  rq_init_comm_if_connected(9, "1")
  rq_init_comm_if_connected(2, "2")
  rq_init_comm_if_connected(3, "3")
  rq_init_comm_if_connected(4, "4")
  rq_print_connected_grippers()
  rq_gripper_communication_thread = run rq_gripper_communication()
  set_closed_norm(97.6470588235294, 1)
  set_open_norm(1.1764705882352942, 1)
  set_closed_mm(0.0, 1)
  set_open_mm(53.0, 1)
  set_closed_norm(100.0, 2)
  set_open_norm(0.0, 2)
  set_closed_mm(0.0, 2)
  set_open_mm(50.0, 2)
  set_closed_norm(100.0, 3)
  set_open_norm(0.0, 3)
  set_closed_mm(0.0, 3)
  set_open_mm(50.0, 3)
  set_closed_norm(100.0, 4)
  set_open_norm(0.0, 4)
  set_closed_mm(0.0, 4)
  set_open_mm(50.0, 4)
  rq_current_limit_enabled = False
  while(not rq_gripper_communication_thread_started):
      sync()
  end
  # end: URCap Installation Node
  # begin: URCap Installation Node
  #   Source: OPC UA, 2.0.2, Rocketfarm AS
  #   Type: OPC UA
  global opcua_daemon = rpc_factory("xmlrpc", "http://127.0.0.1:40409/RPC2")
  def opcua_client_connect(address):
  return opcua_daemon.client_connect(address)
  end
  def opcua_client_get_id(client_name):
  return opcua_daemon.client_get_id(client_name)
  end
  def opcua_client_try_connect(client_id):
  opcua_result = False
  if (opcua_daemon.client_connect(client_id)):
  sleep(0.01)
  opcua_result = opcua_daemon.client_is_connected(client_id)
  opcua_retry = 10
  while ( (not opcua_result) and (opcua_retry > 0) ):
  sleep(0.1)
  opcua_result = opcua_daemon.client_is_connected(client_id)
  opcua_retry = opcua_retry - 1
  end
  end
  return opcua_result
  end
  def opcua_client_disconnect(client_id):
  return opcua_daemon.client_disconnect(client_id)
  end
  def opcua_client_is_connected(client_id):
  return opcua_daemon.client_is_connected(client_id)
  end
  def opcua_client_read_byid(client_id, namespace_id, variable_id):
  return opcua_daemon.client_read_variable_by_id(client_id, namespace_id, variable_id)
  end
  def opcua_client_read_byname(client_id, namespace_id, variable_name):
  return opcua_daemon.client_read_variable_by_name(client_id, namespace_id, variable_name)
  end
  def opcua_client_write_byid(client_id, namespace_id, variable_id, variable_value):
  return opcua_daemon.client_write_variable_by_id(client_id, namespace_id, variable_id, variable_value)
  end
  def opcua_client_write_byname(client_id, namespace_id, variable_name, variable_value):
  return opcua_daemon.client_write_variable_by_name(client_id, namespace_id, variable_name, variable_value)
  end
  def opcua_client_last_error(client_id):
  return opcua_daemon.client_get_last_error(client_id)
  end
  def opcua_server_read_byname(variable_name):
  return opcua_daemon.server_read_variable_by_name(variable_name)
  end
  def opcua_server_write_byname(variable_name, variable_value):
  return opcua_daemon.server_write_variable_by_name(variable_name, variable_value)
  end
  def opcua_server_last_error():
  return opcua_daemon.server_get_last_error()
  end
  def opcua_error_to_string(errorCode):
  return opcua_daemon.error_code_to_string(errorCode)
  end
  # end: URCap Installation Node
  step_count_7f95097d_1581_4d0e_9124_3b7fc3d01574 = 0.0
  thread Step_Counter_Thread_7db62caa_18b4_480e_a8f7_ee898fbd2f33():
    while (True):
      step_count_7f95097d_1581_4d0e_9124_3b7fc3d01574 = step_count_7f95097d_1581_4d0e_9124_3b7fc3d01574 + 1.0
      sync()
    end
  end
  run Step_Counter_Thread_7db62caa_18b4_480e_a8f7_ee898fbd2f33()
  global AMR_Position=struct(position_identifier=0, x1=0, x2=0, y1=0, y2=0, theta1=0, theta2=0)
  global CAM_Pose=p[0,0,0,0,0,0]
  global CAM_Relation=""
  global CMD_Abort=  False
  global CMD_Clear=  False
  global CMD_Reset=  False
  global CMD_Start=  False
  global CMD_Suspend=  False
  global CMD_Unhold=  False
  global CMD_Unsuspend=  False
  global CNT_Rack_Output=0
  global FNC_Freedrive=  False
  global PRC_TubCounter=0
  global PRC_TubNumber=0
  global STP=0
  global easyPickCount=0
  global easyPickCount_5=0
  global easyPickNoObj=0
  global easyPickNoObj_5=0
  global easyPickParts=0
  global easyPickParts_5=0
  global TMR_Barcode=0
  global Container_mid_1_p=p[-.379239199143, -.127191311915, .299999999998, .000000000046, -.000000000021, -1.247199999994]
  global Container_mid_1_q=[-2.477408934449926, -1.2969853503591224, -1.875639182904262, -1.539621866126728, 1.5731943360401213, -2.8009955944022717]
  global Container_capt_p=p[-.525590029047, .407247642794, .411588185841, -.000000000107, .000000000065, -2.896148821900]
  global Container_capt_q=[-3.5968351615224767, -2.0050156108707204, -0.8176271154495112, -1.8895759482008394, 1.5730967555598792, -2.2743681102957645]
  global Waypoint_6_p=p[.008800512419, -.547926542621, .402696567415, -.589884378425, -.007228654778, -.061268144704]
  global Waypoint_6_q=[-1.2044575850116175, -1.3416667741588135, -1.8272563219070435, -0.9884541195682068, 1.3621035814285278, -2.7712565104113978]
  global Waypoint_18_p=p[-.178371829612, -.433927395311, .368082383916, -.086593488055, .704679941724, -.007869906074]
  global Waypoint_18_q=[-1.265390698109762, -1.3355963987163086, -1.7944865226745605, -1.7402602634825648, 0.8780410885810852, -2.7713127771960657]
  global Waypoint_12_p=p[.008800512419, -.547926542621, .402696567415, -.589884378425, -.007228654778, -.061268144704]
  global Waypoint_12_q=[-1.2044575850116175, -1.3416667741588135, -1.8272563219070435, -0.9884541195682068, 1.3621035814285278, -2.7712565104113978]
  global Waypoint_19_p=p[-.178371829612, -.433927395311, .368082383916, -.086593488055, .704679941724, -.007869906074]
  global Waypoint_19_q=[-1.265390698109762, -1.3355963987163086, -1.7944865226745605, -1.7402602634825648, 0.8780410885810852, -2.7713127771960657]
  global Vial_above_p=p[.017105793010, -.652093028359, .184920586844, .000000000272, .000000000270, 1.564063451276]
  global Vial_above_q=[-1.3375440709712851, -1.9618096977868804, -1.4665759083780685, -1.2837941559171444, 1.5732503672317195, -4.47276330421513]
  global Vial_pick_point_p=p[.017105792852, -.648922724010, .093307568731, .000000000271, .000000000270, 1.564063451276]
  global Vial_pick_point_q=[-1.3366329456391917, -2.0375277831965413, -1.6071432798879028, -1.0675084332049813, 1.57309887265915, -4.471135348858068]
  global Waypoint_20_p=p[.019227646885, -.648669633640, .184920586950, .000000000000, .000000000000, .024063451426]
  global Waypoint_20_q=[-1.3331129109407733, -1.9540750545686123, -1.4775914902901128, -1.280581784992414, 1.5733500744865856, -2.928303704452631]
  global Waypoint_33_p=p[-.032361834699, -.348336136197, .391475576335, -.000008499254, .000014589902, -.004651426820]
  global Waypoint_33_q=[-1.2709335019096129, -1.1914598663441005, -1.708995335060501, -1.8117888533498316, 1.5729683532263925, -2.8379347397710237]
  global Vial_3FG_place_p=p[-.031858676359, -.349402499566, .145301120695, .000000000000, .000000000000, .000000000000]
  global Vial_3FG_place_q=[-1.2723975525801707, -1.252376585823825, -2.3128114007049496, -1.1470592278900167, 1.5730548099411423, -2.8414815174610535]
  global Waypoint_34_p=p[-.032361834699, -.348336136197, .391475576335, -.000008499254, .000014589902, -.004651426820]
  global Waypoint_34_q=[-1.2709335019096129, -1.1914598663441005, -1.708995335060501, -1.8117888533498316, 1.5729683532263925, -2.8379347397710237]
  global cap_dump_p=p[-.139168676487, -.420163541420, .146096395183, .000000000000, .000000000000, .000000000000]
  global cap_dump_q=[-1.584588644510994, -1.5093464179777323, -2.1118449369620347, -1.091059703602438, 1.5728943834877336, -3.154014906686923]
  global Waypoint_35_p=p[-.032361834699, -.348336136197, .391475576335, -.000008499254, .000014589902, -.004651426820]
  global Waypoint_35_q=[-1.2709335019096129, -1.1914598663441005, -1.708995335060501, -1.8117888533498316, 1.5729683532263925, -2.8379347397710237]
  global Waypoint_36_p=p[-.032361834699, -.348336136197, .391475576335, -.000008499254, .000014589902, -.004651426820]
  global Waypoint_36_q=[-1.2709335019096129, -1.1914598663441005, -1.708995335060501, -1.8117888533498316, 1.5729683532263925, -2.8379347397710237]
  global Waypoint_37_p=p[-.032361834699, -.348336136197, .391475576335, -.000008499254, .000014589902, -.004651426820]
  global Waypoint_37_q=[-1.2709335019096129, -1.1914598663441005, -1.708995335060501, -1.8117888533498316, 1.5729683532263925, -2.8379347397710237]
  global Vial_liq_above_p=p[-.025303660977, -.338758622354, .426628485936, -1.315858642253, .800043520260, -.928295855026]
  global Vial_liq_above_q=[-0.3789628187762659, -1.5149522957256814, -2.263045310974121, 0.7870649534412841, -0.750984017048971, -3.2237566153155726]
  global Vial_liq_pick_1_p=p[-.002660428945, -.335984893034, .159389832934, -1.150456778400, .673175527684, -1.010612657503]
  global Vial_liq_pick_1_q=[-0.3660772482501429, -1.4503649038127442, -2.4056053161621094, -1.994692941705221, 0.8039668202400208, -0.2508929411517542]
  global Vial_liq_pick_2_p=p[-.041402486291, -.356791603314, .125395323246, -1.143483969075, .651070210027, -.878721885453]
  global Vial_liq_pick_2_q=[-0.4426233705502476, -1.437252121513727, -2.551930962114307, -1.776528229806984, 0.6562026234073748, -0.43018811960029524]
  global Liquid_midway_p=p[.057575295009, -.583081747994, .306414980749, -1.351675548728, .120935756539, -.096908606303]
  global Liquid_midway_q=[-0.895174805318014, -1.7035466633238734, -2.380953073501587, 0.631549521083496, 0.7706599235534668, -2.9455552736865442]
  global shake_1_p=p[.057574880217, -.583085370269, .306422893466, -1.360996190983, -.155555042453, -.438136255921]
  global shake_1_q=[-0.8951800505267542, -1.7035466633238734, -2.380937099456787, 0.6315542894550782, 0.7706599235534669, -2.5394540616517496]
  global shake_2_p=p[.057581636113, -.583090570002, .306439684073, -1.308767904323, .368530312677, .214926493520]
  global shake_2_q=[-0.8951714674579065, -1.7035395107665003, -2.380906343460083, 0.6315504747578125, 0.7706480026245118, -3.3161255787892268]
  global drop_above_1_p=p[.268235025993, -.467784390499, .226219872376, -1.027832627524, -.430841408251, 1.004603115937]
  global drop_above_1_q=[-0.935645882283346, -1.6663371525206507, -2.4252893924713135, 0.41966931402172847, 1.8470635414123535, -3.4600217978106897]
  global drop_above_2_p=p[.219042229014, -.470775657081, .133754190740, -.313004595901, -.344395319364, 1.500564994056]
  global drop_above_2_q=[-1.0601594887284795, -1.70046459045642, -2.0799996233759863, -0.7243227230676759, 1.9429634314685202, -4.115129153870795]
  global liq_tran_1_p=p[.213067510942, -.469567035397, .100231043184, .251862243732, .217902579404, 1.592812335393]
  global liq_tran_1_q=[-0.7789645168037476, -1.822364827406652, -1.8643518410805573, -1.252158963840138, 1.3768134449520435, -3.9328333233290254]
  global Waypoint_21_p=p[.187119460405, -.493959476151, .133754190608, -.313004596540, -.344395317757, 1.500564993991]
  global Waypoint_21_q=[-1.1418328121400876, -1.7310553375189475, -2.033634768766424, -0.772026910513711, 1.958578934631971, -4.201588449364511]
  global liq_tran_2_p=p[.195957706507, -.493022614126, .100231042689, .160718757180, .109807038912, 1.525321508623]
  global liq_tran_2_q=[-0.881740380645474, -1.8244526267589851, -1.865100964490387, -1.1608866323693583, 1.4631433601076713, -3.973915130363038]
  global Vial_drop_above_p=p[.000324902251, -.648569523142, .221894115667, -.873462921366, 1.165852672573, -1.482720593185]
  global Vial_drop_above_q=[-1.0576906334721352, -2.393016994184633, -0.9236232851859159, -2.5729213042279273, 0.7903331288549689, -0.33286325848155585]
  global Vial_liq_drop_p=p[.001020867953, -.647659915585, .092915870838, -.834762611599, 1.081942994823, -1.540647900176]
  global Vial_liq_drop_q=[-1.0631954168193474, -2.4447642951220825, -1.128811017825127, -2.1983115491972294, 0.8130148661460634, -0.38984988696911316]
  global Waypoint_9_p=p[.206300564882, -.401796282405, .209941275233, .000000000049, .000000000063, 1.560839127857]
  global Waypoint_9_q=[-0.7963359454512808, -1.4686025034365713, -1.9726632321075135, -1.2709582822971974, 1.5730203818053559, -3.9272300959189193]
  global Waypoint_10_p=p[.200865824304, -.400817692024, .105072686738, .000000000049, .000000000061, 1.560839127855]
  global Waypoint_10_q=[-0.8042914374275529, -1.5824702465090397, -2.1630314773482997, -0.9667217216455377, 1.5726337265768082, -3.9342465798801403]
  global Waypoint_11_p=p[.200865824280, -.400817691999, .325177251663, .000000000049, .000000000061, 1.560839127855]
  global Waypoint_11_q=[-0.8031609769098491, -1.4190566846320642, -1.7173307870816634, -1.5758364190022327, 1.5730457436482617, -3.935202548332848]
  global Waypoint_7_p=p[-.615828862681, .233809157513, .299999999960, .005115849907, .008741794022, -2.111813105778]
  global Waypoint_7_q=[-3.2957401409809868, -1.9361965884744503, -1.2056078493731617, -1.569266158150004, 1.5650998100608482, -2.7562028470627613]
  global Waypoint_8_p=p[-.615828862366, .233809157463, .013910424379, .005115849905, .008741794020, -2.111813105780]
  global Waypoint_8_q=[-3.2964782505943173, -2.1586184138220776, -1.6500090431308791, -0.9024541777239836, 1.5648120752692236, -2.7547026290098384]
  global Waypoint_13_p=p[-.479450777041, .284140798427, .125270103493, -.276792173670, 2.098433187455, -2.121256516887]
  global Waypoint_13_q=[-2.8915050665484827, -1.9549266300597132, -2.2318272590637207, -1.6654960117735804, 0.020810842514038086, -0.4019392172442835]
  global Waypoint_70_p=p[-.472820924464, .292439826304, .207418370234, -.259787347864, -2.053484648504, 2.070709755662]
  global Waypoint_70_q=[-2.969927421603815, -2.07168115810532, -1.6835546062719366, -2.4953958198513964, 0.4489790927922641, -0.005578998612037367]
  global Waypoint_1_p=p[-.312961047461, -.152991312519, .223609826854, -.745314530454, -1.713873240489, 1.673341715282]
  global Waypoint_1_q=[-2.3560472170459192, -2.183784624139303, -1.4583134651184082, -2.6435262165465296, 1.6522362232208252, 0.043451953679323196]
  global Waypoint_16_p=p[-.113749865836, -.390110151572, .317307487562, -.519383711706, -.839884211339, 1.756868173041]
  global Waypoint_16_q=[-1.8909733931170862, -1.720626016656393, -1.5115610361099243, -2.1240560017027796, 2.1809096336364746, 0.7227501273155212]
  global Waypoint_15_p=p[.029144035010, -.436802470887, .327885032028, -.521560953301, -.623641814548, 1.862659450154]
  global Waypoint_15_q=[-1.564817253743307, -1.556895188321807, -1.6826975345611572, -1.6944714985289515, 2.2362685203552246, 1.117417335510254]
  global Waypoint_14_p=p[.068712235638, -.569419545175, .285215357659, -.679242949116, -.712065334485, 1.394044574094]
  global Waypoint_14_q=[-1.5731792953485346, -1.8029235103747094, -1.6781008808776736, -1.2218450646111982, 2.4719572998240125, 1.6394218026856375]
  global Waypoint_17_p=p[-.047220457210, -.557624911767, .136370962514, -.679242949107, -.712065334475, 1.394044574096]
  global Waypoint_17_q=[-1.7740079055958748, -2.0023561428872334, -1.7577251142892676, -1.18903287716154, 2.4487287370345143, 1.322902469273079]
  global Waypoint_25_p=p[.065436479647, -.569388431626, .287820755049, -.679242949185, -.712065334557, 1.394044574070]
  global Waypoint_25_q=[-1.5789263550890595, -1.8020194754825436, -1.6702557537748035, -1.237882536889547, 2.471995808083492, 1.6301087487321393]
  global Waypoint_73_p=p[.200650292861, -.570238752026, .330084459991, 1.360500825815, .021700154388, 2.681649888469]
  global Waypoint_73_q=[-0.7671117850166942, -2.170180210127774, -0.8654875324671831, -2.4760661058854714, 1.019668964673781, 1.1886838746103445]
  global Waypoint_51_p=p[.143029822311, -.569853361759, .275754213782, 1.297896664289, .026410127072, 2.712872144875]
  global Waypoint_51_q=[-0.8339941389801577, -2.0499669090260237, -1.181859109742545, -2.1992567984298894, 0.9933974691724003, 1.1053015960835664]
  global Waypoint_55_p=p[.073857253409, -.577012553496, .221504790513, 1.297896665457, .026410123899, 2.712872144362]
  global Waypoint_55_q=[-0.9235026509638331, -2.0031911550113533, -1.4013130080059835, -1.9791459123699324, 0.9364696407276547, 1.0224867664664226]
  global Waypoint_56_p=p[.135677267144, -.579447716527, .242231366835, 1.555421348248, .015405426287, 2.555899922373]
  global Waypoint_56_q=[-0.8277598345563266, -2.1783820448240228, -1.1390951780517948, -2.3437042464770936, 0.9222576608739947, 1.2572681804986878]
  global Waypoint_57_p=p[.143391004007, -.581808738942, .226065325532, 1.639743959545, .007914821713, 2.502360786858]
  global Waypoint_57_q=[-0.8163397121067408, -2.2409861865625498, -1.1056400409378426, -2.4000192569642436, 0.9131014133193622, 1.3141118037187605]
  global Waypoint_59_p=p[.272401132286, -.578182925380, .239561357365, 2.126997331910, .113921148153, 2.155615020515]
  global Waypoint_59_q=[-0.6600120703326624, -2.700596948663229, -0.4450863301753998, -3.1158048115172328, 0.9327830672264099, 1.686402678489685]
  global Waypoint_58_p=p[.223648508176, -.578477552733, .276546452136, 2.174288010107, -.044108754041, 2.058653287678]
  global Waypoint_58_q=[-0.7290484882560344, -2.6749849159411134, -0.44426632073579775, -3.220833992584847, 0.9665895014735898, 1.686536774549042]
  global Waypoint_60_p=p[-.013316432876, -.544772031582, .383371643081, 2.208233379808, .037543335712, 2.097559881761]
  global Waypoint_60_q=[-0.9328326161883087, -2.0999933666355775, -1.1958015693111372, -3.060905141293654, 0.690378518537611, 1.7121940951337198]
  global Waypoint_61_p=p[-.412188693372, -.356446875193, .383371643081, 1.751740964455, -.739956256289, 1.600691174920]
  global Waypoint_61_q=[-1.766185342973321, -2.0999933666355775, -1.1958015693111372, -3.060905141293654, 0.690378518537611, 1.7121940951337198]
  global Waypoint_62_p=p[-.542658707241, -.114281911009, .251261544113, 1.813043609523, -.679411528034, 1.655271622964]
  global Waypoint_62_q=[-2.158300033470912, -1.9418836862428677, -1.8142999147147894, -2.778920736683023, 0.21900622104017292, 1.8983390235012934]
  global Waypoint_63_p=p[-.532496162227, -.127810170801, .159342327524, 1.813043609478, -.679411528027, 1.655271622994]
  global Waypoint_63_q=[-2.1232624524640213, -2.086114053133292, -1.8911847933380095, -2.5248779786918614, 0.2536249317365024, 1.864405460969639]
  global Waypoint_52_p=p[-.576034890047, -.066269986912, .306739617770, .862065193359, -.255405331227, 2.195240951653]
  global Waypoint_52_q=[-2.4808268779922003, -1.5303848711262056, -1.876845562237385, -1.1257011427858359, 0.8740163290385958, -0.15002503295170655]
  global Waypoint_69_p=p[-.581965326699, -.059291422286, .312082125679, .862065195757, -.255405329473, 2.195240950921]
  global Waypoint_69_q=[-2.500621389999687, -1.5361955180345959, -1.8614018767844556, -1.1190332887072278, 0.8777181708365909, -0.17540933674578696]
  global Waypoint_71_p=p[-.581965326670, -.059291422265, .290575803625, .862065195756, -.255405329472, 2.195240950921]
  global Waypoint_71_q=[-2.5007210652259566, -1.5510704265538795, -1.9040561970342402, -1.0615823481403304, 0.8776641555740685, -0.17528706367848557]
  global Waypoint_72_p=p[-.581965326627, -.059291422244, .350142125738, 1.757497900770, -.677813691618, 1.696469016977]
  global Waypoint_72_q=[-2.3014470577960933, -1.774776476208789, -1.7081605706825291, -2.8433626113276596, 0.07508598567825443, 1.682946898281932]
  global Waypoint_68_p=p[-.333292906431, -.480744165508, .350142125738, 2.217519979286, .140864133573, 2.209123277630]
  global Waypoint_68_q=[-1.438387057796029, -1.774776476208789, -1.7081605706825291, -2.8433626113276596, 0.07508598567825443, 1.682946898281932]
  global TMR_Barcode_is_counting=False
  thread Timer_Thread():
    while (True):
      if (TMR_Barcode_is_counting):
        TMR_Barcode = TMR_Barcode + get_steptime()
      end
      sync()
    end
  end
  run Timer_Thread()
  def Sub_Vision_V18():
    $ 882 "Sub_Vision_V18" "noBreak"
    $ 883 "PreSettings"
    $ 884 "CAM_LM_Detected≔ False "
    global CAM_LM_Detected=  False
    $ 885 "CAM_Captures≔0"
    global CAM_Captures=0
    $ 886 "CAM_Pose≔p[0,0,0,0,0,0]"
    global CAM_Pose=p[0,0,0,0,0,0]
    $ 887 "CAM_LM_Refinmnt≔ False "
    global CAM_LM_Refinmnt=  False
    $ 888 "CAM_LM_Refined≔ False "
    global CAM_LM_Refined=  False
    $ 889 "CAM_LM_Deviatn≔p[0,0,0,0,0,0]"
    global CAM_LM_Deviatn=p[0,0,0,0,0,0]
    $ 890 "CAM_LM_ID≔0"
    global CAM_LM_ID=0
    $ 891 "CAM_Done≔ False "
    global CAM_Done=  False
    $ 892 "CAM_CNT_Obj≔0"
    global CAM_CNT_Obj=0
    $ 893 "CAM_Result = []"
    CAM_Result = []
    $ 894 "OBJ_Detected≔ False "
    global OBJ_Detected=  False
    $ 895 "FRM_Reference≔p[0,0,0,0,0,0]"
    global FRM_Reference=p[0,0,0,0,0,0]
    $ 896 "'=========='"
    # '=========='
    $ 897 "Switch Action"
    switch_1 = Action
    $ 898 "Case 13"
    if (13 == switch_1):
    elif (15 == switch_1):
      $ 1016 "Case 15"
    elif (131 == switch_1):
      $ 1062 "Case 131"
      $ 1063 "Read (SensoPart)"
      $ 1064 "Action_Info≔'search for landmark'"
      global Action_Info="search for landmark"
      $ 1065 "CAM_LM≔CAM_LMs[4]"
      global CAM_LM=CAM_LMs[4]
      $ 1066 "CAM_Relation≔CAM_LM.capture_relation"
      global CAM_Relation=CAM_LM.capture_relation
      $ 1067 "go to capture pose"
      $ 1070 "If ITM_ID≟1 and JIG≟7"
      if (ITM_ID == 1  and  JIG == 7):
        $ 1071 "PSE_T≔uLM_Cap_SSRack"
        global PSE_T=uLM_Cap_SSRack
      else:
        $ 1072 "ElseIf ITM_ID≟5 and JIG≟7"
        if (ITM_ID == 5  and  JIG == 7):
          $ 1073 "PSE_T≔FRM_Cap_SSRack"
          global PSE_T=FRM_Cap_SSRack
        else:
          $ 1074 "ElseIf ITM_ID≟13 and JIG≟7"
          if (ITM_ID == 13  and  JIG == 7):
            $ 1075 "PSE_T≔FRM_pick_rack_const"
            global PSE_T=p[0.0,0.0,0.0,0.0,0.0,0.0]
          else:
            $ 1076 "ElseIf ITM_ID≟1 and JIG≟15"
            if (ITM_ID == 1 and JIG == 15):
              $ 1077 "MoveJ"
              $ 1078 "Container_mid_1" "breakAfter"
              movej(get_inverse_kin(Container_mid_1_p, qnear=Container_mid_1_q), a=1.3962634015954636, v=1.0471975511965976, r=0.05)
              $ 1079 "Container_capt" "breakAfter"
              movej(get_inverse_kin(Container_capt_p, qnear=Container_capt_q), a=1.3962634015954636, v=1.0471975511965976)
              $ 1080 "PSE_T≔FRM_Container_S_const"
              global PSE_T=p[0.0,0.0,0.0,0.0,0.0,0.0]
            end
          end
        end
      end
      $ 1081 "do_transition(PSE_T, keep_rxry=False)"
      do_transition(PSE_T, keep_rxry=False)
      $ 1082 "Set"
      set_tcp(p[0.0,0.0,0.161,3.1415,0.0,0.0])
      $ 1083 "MoveJ"
      $ 1084 "PSE_T" "breakAfter"
      movej(PSE_T, a=1.3962634015954636, v=1.7453292519943295)
      $ 1085 "CAM_Pose≔get_actual_tcp_pose()"
      global CAM_Pose= get_actual_tcp_pose ()
      $ 1086 "Loop  not CAM_Done and  not ERROR.FLAG and  not CMD_Stop"
      while (  not  CAM_Done  and    not  ERROR.FLAG  and    not  CMD_Stop):
        $ 1087 "adjust capture pose"
        $ 1088 "If CAM_LM_Detected and CAM_LM_Refinmnt"
        if (CAM_LM_Detected  and  CAM_LM_Refinmnt):
          $ 1089 "PSE_T≔p[0,0,0.300,0,0,0]"
          global PSE_T=p[0,0,0.300,0,0,0]
          $ 1090 "CAM_Pose≔PSE_T"
          global CAM_Pose=PSE_T
          $ 1091 "If  not is_reachable(FRM_Reference,[PSE_T])"
          if (  not  is_reachable(FRM_Reference,[PSE_T])):
            $ 1092 "Error"
            $ 1093 "set_error(ERROR_POSE_NOT_REACHABLE)"
            set_error(ERROR_POSE_NOT_REACHABLE)
          end
          $ 1094 "If  not ERROR.FLAG"
          if (  not  ERROR.FLAG):
            $ 1095 "MoveJ"
            $ 1096 "PSE_T" "breakAfter"
            set_tcp(p[0.0,0.0,0.161,0.0,0.0,0.0])
            movej(pose_trans(FRM_Reference, PSE_T), a=0.8726646259971648, v=1.3962634015954636)
            $ 1097 "CAM_LM_Refined≔ True "
            global CAM_LM_Refined=  True
          end
        else:
          $ 1098 "ElseIf  not CAM_LM_Detected and CAM_Captures>0"
          if (  not  CAM_LM_Detected  and  CAM_Captures>0):
            $ 1099 "MoveL"
            $ 1100 "If FRM_Reference≟p[0,0,0,0,0,0]"
            if (FRM_Reference == p[0,0,0,0,0,0]):
              $ 1101 "PSE_T≔get_random_pose(pose_ref=CAM_Pose, mode='cubic', range_max=[0.150,0.150,0.015])"
              global PSE_T=get_random_pose(pose_ref=CAM_Pose, mode="cubic", range_max=[0.150,0.150,0.015])
            else:
              $ 1106 "Else" "noBreak"
              $ 1107 "PSE_T≔get_random_pose(pose_ref=CAM_Pose, mode='rotation', range_max=[10,10,0])"
              global PSE_T=get_random_pose(pose_ref=CAM_Pose, mode="rotation", range_max=[10,10,0])
              $ 1108 "CAM_LM_Refined≔ True "
              global CAM_LM_Refined=  True
            end
            $ 1109 "If get_inverse_kin_has_solution(pose_trans(FRM_Reference, PSE_T))"
            if (get_inverse_kin_has_solution( pose_trans (FRM_Reference, PSE_T))):
              $ 1110 "Comment"
              # Comment
              $ 1111 "PSE_T" "breakAfter"
              set_tcp(p[0.0,0.0,0.161,3.1415,0.0,0.0])
              movel(pose_trans(FRM_Reference, PSE_T), a=0.03, v=0.05)
            else:
              $ 1112 "Else" "noBreak"
              $ 1113 "'If random pose is out of reach, set the initial cam pose'"
              # 'If random pose is out of reach, set the initial cam pose'
              $ 1114 "PSE_T≔CAM_Pose"
              global PSE_T=CAM_Pose
            end
          end
        end
        $ 1115 "Wait: 2.0"
        sleep(2.0)
        $ 1116 "trigger"
        $ 1117 "If ITM_ID≟1 and JIG≟7"
        if (ITM_ID == 1  and  JIG == 7):
          # begin: URCap Program Node
          #   Source: SensoPart VISOR Robotic, 2.0.0, SensoPart Industriesensorik GmbH
          #   Type: VISOR Trigger
          $ 1118 "# 1 VISOR Trigger"
          visor_changeJob(1, "Landmark_INVITE_2", 6000)
          visor_trigger(1, 6000, "arm")
          # end: URCap Program Node
        else:
          $ 1119 "ElseIf ITM_ID≟5 and JIG≟7"
          if (ITM_ID == 5  and  JIG == 7):
            # begin: URCap Program Node
            #   Source: SensoPart VISOR Robotic, 2.0.0, SensoPart Industriesensorik GmbH
            #   Type: VISOR Trigger
            $ 1120 "# 1 VISOR Trigger"
            visor_changeJob(1, "Landmark_INVITE_2", 6000)
            visor_trigger(1, 6000, "arm")
            # end: URCap Program Node
          else:
            $ 1121 "ElseIf ITM_ID≟13 and JIG≟7"
            if (ITM_ID == 13  and  JIG == 7):
              # begin: URCap Program Node
              #   Source: SensoPart VISOR Robotic, 2.0.0, SensoPart Industriesensorik GmbH
              #   Type: VISOR Trigger
              $ 1122 "# 1 VISOR Trigger"
              visor_changeJob(1, "Landmark_INVITE_2", 6000)
              visor_trigger(1, 6000, "arm")
              # end: URCap Program Node
            else:
              $ 1123 "ElseIf ITM_ID≟1 and JIG≟15"
              if (ITM_ID == 1 and JIG == 15):
                # begin: URCap Program Node
                #   Source: SensoPart VISOR Robotic, 2.0.0, SensoPart Industriesensorik GmbH
                #   Type: VISOR Trigger
                $ 1124 "# 1 VISOR Trigger"
                visor_changeJob(1, "Container_S", 6000)
                visor_trigger(1, 6000, "arm")
                # end: URCap Program Node
              end
            end
          end
        end
        $ 1128 "TM_3D_Found≔visor_partsFound(1)"
        global TM_3D_Found= visor_partsFound (1)
        $ 1129 "If TM_3D_Found>0"
        if (TM_3D_Found>0):
          $ 1130 "CAM_LM_Detected≔ True "
          global CAM_LM_Detected=  True
          $ 1131 "CAM_Captures≔0"
          global CAM_Captures=0
        else:
          $ 1132 "Else" "noBreak"
          $ 1133 "CAM_LM_Detected≔ False "
          global CAM_LM_Detected=  False
          $ 1134 "CAM_Captures≔CAM_Captures+1"
          global CAM_Captures=CAM_Captures+1
        end
        $ 1139 "result"
        $ 1140 "If CAM_LM_Detected"
        if (CAM_LM_Detected):
          $ 1141 "If (CAM_LM_Refinmnt and CAM_LM_Refined) or  not CAM_LM_Refinmnt"
          if ((CAM_LM_Refinmnt  and  CAM_LM_Refined)  or    not  CAM_LM_Refinmnt):
            $ 1199 "If ITM_ID≟1 and JIG≟7"
            if (ITM_ID == 1  and  JIG == 7):
              $ 1200 "CAM_LM_SSRack≔visor_getPose3d(1, 0)"
              global CAM_LM_SSRack= visor_getPose3d (1, 0)
            else:
              $ 1201 "ElseIf ITM_ID≟5 and JIG≟7"
              if (ITM_ID == 5  and  JIG == 7):
                $ 1202 "CAM_LM_SSRack≔visor_getPose3d(1, 0)"
                global CAM_LM_SSRack= visor_getPose3d (1, 0)
              end
            end
            $ 1207 "CAM_Done≔ True "
            global CAM_Done=  True
          end
        else:
          $ 1208 "ElseIf  not CAM_LM_Detected and CAM_Captures<CAM_PRM_Retries"
          if (  not  CAM_LM_Detected  and  CAM_Captures<CAM_PRM_Retries):
            $ 1209 "CAM_LM_Refined≔ False "
            global CAM_LM_Refined=  False
          else:
            $ 1210 "ElseIf CAM_Captures≥CAM_PRM_Retries"
            if (CAM_Captures >= CAM_PRM_Retries):
              $ 1211 "CAM_Done≔ True "
              global CAM_Done=  True
              $ 1212 "Error"
              $ 1213 "set_error(ERROR_NO_LANDMARK)"
              set_error(ERROR_NO_LANDMARK)
            end
          end
        end
      end
    elif (151 == switch_1):
      $ 1214 "Case 151"
      $ 1215 "Detect (SensoPart)"
      $ 1216 "go to capture pose"
      $ 1217 "FRM_Reference≔FRM_Cap_SSRack"
      global FRM_Reference=FRM_Cap_SSRack
      $ 1218 "PSE_T≔p[0,0,-0.00,0,0,0]"
      global PSE_T=p[0,0,-0.00,0,0,0]
      $ 1219 "do_transition(pose_trans(FRM_Reference, PSE_T), keep_rxry=False)"
      do_transition( pose_trans (FRM_Reference, PSE_T), keep_rxry=False)
      $ 1220 "JNT_Q≔get_actual_joint_positions()"
      global JNT_Q= get_actual_joint_positions ()
      $ 1221 "JNT_Q≔[JNT_Q[0], JNT_Q[1], JNT_Q[2], JNT_Q[3], JNT_Q[4], 0]"
      global JNT_Q=[JNT_Q[0], JNT_Q[1], JNT_Q[2], JNT_Q[3], JNT_Q[4], 0]
      $ 1222 "Set"
      set_tcp(p[0.0,0.0,0.161,3.1415,0.0,0.0])
      $ 1223 "movej(get_inverse_kin(pose_trans(FRM_Reference, PSE_T), qnear=JNT_Q))"
      movej(get_inverse_kin( pose_trans (FRM_Reference, PSE_T), qnear=JNT_Q))
      $ 1224 "CAM_Pose≔pose_trans(pose_inv(FRM_Reference), get_actual_tcp_pose())"
      global CAM_Pose= pose_trans ( pose_inv (FRM_Reference),  get_actual_tcp_pose ())
      $ 1225 "Loop  not CAM_Done and  not ERROR.FLAG and  not CMD_Stop"
      while (  not  CAM_Done  and    not  ERROR.FLAG  and    not  CMD_Stop):
        $ 1226 "If  not OBJ_Detected and CAM_Captures>0"
        if (  not  OBJ_Detected  and  CAM_Captures>0):
          $ 1227 "MoveL"
          $ 1228 "If FRM_Reference≟p[0,0,0,0,0,0]"
          if (FRM_Reference == p[0,0,0,0,0,0]):
            $ 1230 "PSE_T≔get_random_pose(pose_ref=CAM_Pose, mode='rotation', range_max=[15,15,0])"
            global PSE_T=get_random_pose(pose_ref=CAM_Pose, mode="rotation", range_max=[15,15,0])
          else:
            $ 1231 "Else" "noBreak"
            $ 1232 "PSE_T≔get_random_pose(pose_ref=CAM_Pose, mode='rotation', range_max=[10,10,0])"
            global PSE_T=get_random_pose(pose_ref=CAM_Pose, mode="rotation", range_max=[10,10,0])
          end
          $ 1233 "If get_inverse_kin_has_solution(pose_trans(FRM_Reference, PSE_T))"
          if (get_inverse_kin_has_solution( pose_trans (FRM_Reference, PSE_T))):
            $ 1234 "PSE_T" "breakAfter"
            set_tcp(p[0.0,0.0,0.161,3.1415,0.0,0.0])
            movel(pose_trans(FRM_Reference, PSE_T), a=0.03, v=0.05)
          else:
            $ 1235 "Else" "noBreak"
            $ 1236 "'If random pose is out of reach, set the initial cam pose'"
            # 'If random pose is out of reach, set the initial cam pose'
            $ 1237 "PSE_T≔CAM_Pose"
            global PSE_T=CAM_Pose
            $ 1238 "PSE_T" "breakAfter"
            set_tcp(p[0.0,0.0,0.161,3.1415,0.0,0.0])
            movel(pose_trans(FRM_Reference, PSE_T), a=0.03, v=0.05)
          end
        end
        $ 1239 "Wait: 0.5"
        sleep(0.5)
        $ 1240 "Set"
        set_tcp(p[0.0,0.0,0.161,3.1415,0.0,0.0])
        # begin: URCap Program Node
        #   Source: SensoPart VISOR Robotic, 2.0.0, SensoPart Industriesensorik GmbH
        #   Type: VISOR Trigger
        $ 1241 "# 1 VISOR Trigger"
        visor_changeJob(1, "Object Detection Single", 6000)
        visor_trigger(1, 6000, "arm")
        # end: URCap Program Node
        $ 1242 "If visor_isResponseOk(1)"
        if ( visor_isResponseOk (1)):
          $ 1243 "CAM_CNT_Obj≔visor_partsFound(1)"
          global CAM_CNT_Obj= visor_partsFound (1)
          $ 1244 "CAM_OBJ_Pose≔visor_getPose3d(1, 0)"
          global CAM_OBJ_Pose= visor_getPose3d (1, 0)
          $ 1245 "If CAM_CNT_Obj>0"
          if (CAM_CNT_Obj>0):
            $ 1246 "CAM_OBJ_Color≔visor_getAdditionalData(1, 0)"
            global CAM_OBJ_Color= visor_getAdditionalData (1, 0)
            $ 1247 "CAM_DetectScore≔to_num(visor_getAdditionalData(1, 1))/1000"
            global CAM_DetectScore=to_num( visor_getAdditionalData (1, 1))/1000
            $ 1248 "OBJ_Detected≔ True "
            global OBJ_Detected=  True
          end
        else:
          $ 1249 "Else" "noBreak"
          $ 1250 "CAM_Captures≔CAM_Captures+1"
          global CAM_Captures=CAM_Captures+1
        end
        $ 1251 "If OBJ_Detected"
        if (OBJ_Detected):
          $ 1252 "Get object data"
          $ 1253 "PRC_CntDetect≔0"
          global PRC_CntDetect=0
          $ 1254 "Loop PRC_CntDetect<CAM_CNT_Obj"
          while (PRC_CntDetect<CAM_CNT_Obj):
            $ 1255 "get object and jig number"
            $ 1256 "If ITM_ID≟1 and JIG≟7"
            if (ITM_ID == 1  and  JIG == 7):
              $ 1257 "FRM_Reference≔FRM_Cap_SSRack"
              global FRM_Reference=FRM_Cap_SSRack
            else:
              $ 1258 "ElseIf ITM_ID≟5 and JIG≟7"
              if (ITM_ID == 5  and  JIG == 7):
                $ 1259 "FRM_Reference≔uLM_Cap_SSRack"
                global FRM_Reference=uLM_Cap_SSRack
              end
            end
            $ 1262 "PSE_T≔pose_trans(pose_inv(FRM_Reference), CAM_OBJ_Pose)"
            global PSE_T= pose_trans ( pose_inv (FRM_Reference), CAM_OBJ_Pose)
            $ 1263 "CAM_Result.append(get_pattern_counter(PSE_T, 'X', pattern=[10, 5], patternsize=[0.181, 0.081]))"
            CAM_Result.append(get_pattern_counter(PSE_T, "X", pattern=[10, 5], patternsize=[0.181, 0.081]))
            $ 1264 "PRC_CntDetect≔PRC_CntDetect+1"
            global PRC_CntDetect=PRC_CntDetect+1
          end
          $ 1265 "CAM_Done≔ True "
          global CAM_Done=  True
        else:
          $ 1266 "ElseIf CAM_Captures≥CAM_PRM_Retries"
          if (CAM_Captures >= CAM_PRM_Retries):
            $ 1267 "CAM_Done≔ True "
            global CAM_Done=  True
          else:
            $ 1268 "Else" "noBreak"
            $ 1269 "CAM_Captures≔CAM_Captures+1"
            global CAM_Captures=CAM_Captures+1
          end
        end
      end
    end
    $ 1270 "'=========='"
    # '=========='
    $ 1271 "PostSettings"
    $ 1272 "FRM_Reference≔p[0,0,0,0,0,0]"
    global FRM_Reference=p[0,0,0,0,0,0]
    $ 1273 "Set"
    set_tcp(p[0.0,0.0,0.161,3.1415,0.0,0.0])
    $ 1274 "CAM_Pose≔p[0,0,0,0,0,0]"
    global CAM_Pose=p[0,0,0,0,0,0]
    $ 1275 "Action≔0"
    global Action=0
    $ 1276 "Action_Info≔''"
    global Action_Info=""
  end
  def Sub_AMR_MiR_V3():
    $ 1277 "Sub_AMR_MiR_V3" "noBreak"
    $ 1278 "PreSettings"
    $ 1279 "AMR_TargetList≔[1,2,3,4,5,21,22,23,24,31,32,33,34,35,36,37,38,41]"
    global AMR_TargetList=[1,2,3,4,5,21,22,23,24,31,32,33,34,35,36,37,38,41]
    $ 1280 "AMR_Done≔ False "
    global AMR_Done=  False
    $ 1281 "AMR_PosActual≔T2O_Current_Pos"
    global AMR_PosActual=modbus_get_signal_status("T2O_Current_Pos")
    $ 1282 "AMR_Attemps≔T2O_Nav_Attemps"
    global AMR_Attemps=modbus_get_signal_status("T2O_Nav_Attemps")
    $ 1283 "AMR_Battery≔MiR_Battery_Lvl"
    global AMR_Battery=modbus_get_signal_status("MiR_Battery_Lvl")
    $ 1284 "AMR_Charging≔(T2O_Charging≟1)"
    global AMR_Charging=(modbus_get_signal_status("T2O_Charging") == 1)
    $ 1285 "AMR_Position≔struct(position_identifier=T2O_Current_Pos, x1=MiR_Position_X1, x2=MiR_Position_X2, y1=MiR_Position_Y1, y2=MiR_Position_Y2, theta1=MiR_Theta_1, theta2=MiR_Theta_2) "
    global AMR_Position=struct(position_identifier=modbus_get_signal_status("T2O_Current_Pos"), x1=modbus_get_signal_status("MiR_Position_X1"), x2=modbus_get_signal_status("MiR_Position_X2"), y1=modbus_get_signal_status("MiR_Position_Y1"), y2=modbus_get_signal_status("MiR_Position_Y2"), theta1=modbus_get_signal_status("MiR_Theta_1"), theta2=modbus_get_signal_status("MiR_Theta_2"))
    $ 1286 "If MiR_Mode≠7"
    if (modbus_get_signal_status("MiR_Mode") != 7):
      $ 1287 "Error"
      $ 1288 "set_error(ERROR_AMR_WRONG_MODE)"
      set_error(ERROR_AMR_WRONG_MODE)
      $ 1289 "AMR_Done≔ True "
      global AMR_Done=  True
    end
    $ 1290 "'=========='"
    # '=========='
    $ 1291 "Switch STATE"
    switch_1 = STATE
    $ 1292 "Case 1"
    if (1 == switch_1):
      $ 1293 "stopping"
      $ 1294 "If T2O_Done≟1 and O2T_Acknowledge≟0"
      if (modbus_get_signal_status("T2O_Done") == 1  and  modbus_get_signal_status("O2T_Acknowledge") == 0):
        $ 1295 "Set O2T_Acknowledge=1"
        modbus_set_output_register("O2T_Acknowledge", 1)
      end
      $ 1296 "Set MiR_CMD_Stop=On"
      modbus_set_output_signal("MiR_CMD_Stop", True)
      $ 1297 "AMR_Position.position_identifier = 0"
      AMR_Position.position_identifier = 0
      $ 1298 "AMR_Done≔ True "
      global AMR_Done=  True
    elif (2 == switch_1):
      $ 1299 "Case 2"
      $ 1300 "stopped"
      $ 1301 "If MiR_State≠3 and MiR_State≠5"
      if (modbus_get_signal_status("MiR_State") != 3  and  modbus_get_signal_status("MiR_State") != 5):
        $ 1302 "Set MiR_CMD_Stop=Off"
        modbus_set_output_signal("MiR_CMD_Stop", False)
      end
    elif (3 == switch_1):
      $ 1303 "Case 3"
      $ 1304 "resetting"
      $ 1305 "Set O2T_Mis_Main=Off"
      modbus_set_output_signal("O2T_Mis_Main", False)
      $ 1306 "Set O2T_Mis_Charge=Off"
      modbus_set_output_signal("O2T_Mis_Charge", False)
      $ 1307 "If MiR_Mis_Queue>0"
      if (modbus_get_signal_status("MiR_Mis_Queue")>0):
        $ 1308 "Set MiR_CMD_Clear_Q=On"
        modbus_set_output_signal("MiR_CMD_Clear_Q", True)
        $ 1309 "Wait MiR_Mis_Queue≟0"
        while (not(modbus_get_signal_status("MiR_Mis_Queue") == 0)):
          sync()
        end
        $ 1310 "Set MiR_CMD_Clear_Q=Off"
        modbus_set_output_signal("MiR_CMD_Clear_Q", False)
      end
      $ 1311 "If MiR_Error_ID≠0"
      if (modbus_get_signal_status("MiR_Error_ID") != 0):
        $ 1312 "Set MiR_CMD_Clear_E=On"
        modbus_set_output_signal("MiR_CMD_Clear_E", True)
        $ 1313 "Wait MiR_Error_ID≟0"
        while (not(modbus_get_signal_status("MiR_Error_ID") == 0)):
          sync()
        end
        $ 1314 "Set MiR_CMD_Clear_E=Off"
        modbus_set_output_signal("MiR_CMD_Clear_E", False)
      end
      $ 1315 "Set O2T_Action=0"
      modbus_set_output_register("O2T_Action", 0)
      $ 1316 "Set O2T_Acknowledge=0"
      modbus_set_output_register("O2T_Acknowledge", 0)
      $ 1317 "Set O2T_Target_Pos=0"
      modbus_set_output_register("O2T_Target_Pos", 0)
      $ 1318 "Set O2T_Footprint=0"
      modbus_set_output_register("O2T_Footprint", 0)
      $ 1319 "Set O2T_ProtectOff=0"
      modbus_set_output_register("O2T_ProtectOff", 0)
      $ 1320 "Set O2T_Dock=0"
      modbus_set_output_register("O2T_Dock", 0)
      $ 1321 "AMR_Attemps≔0"
      global AMR_Attemps=0
      $ 1322 "AMR_PosTarget≔0"
      global AMR_PosTarget=0
      $ 1323 "AMR_Step≔0"
      global AMR_Step=0
      $ 1324 "AMR_AtTarget≔ False "
      global AMR_AtTarget=  False
      $ 1325 "If MiR_State≟4 or MiR_State≟3 or MiR_State≟10"
      if (modbus_get_signal_status("MiR_State") == 4  or  modbus_get_signal_status("MiR_State") == 3  or  modbus_get_signal_status("MiR_State") == 10):
        $ 1326 "AMR_Done≔ True "
        global AMR_Done=  True
      end
    elif (5 == switch_1):
      $ 1327 "Case 5"
      $ 1328 "starting"
      $ 1329 "If MiR_State≟4"
      if (modbus_get_signal_status("MiR_State") == 4):
        $ 1330 "Set MiR_CMD_Start=On"
        modbus_set_output_signal("MiR_CMD_Start", True)
        $ 1331 "Wait MiR_State≠4"
        while (not(modbus_get_signal_status("MiR_State") != 4)):
          sync()
        end
        $ 1332 "Set MiR_CMD_Start=Off"
        modbus_set_output_signal("MiR_CMD_Start", False)
        $ 1333 "AMR_Done≔ True "
        global AMR_Done=  True
      else:
        $ 1334 "ElseIf MiR_State≟10"
        if (modbus_get_signal_status("MiR_State") == 10):
          $ 1335 "'MiR in protective stop. Wait'"
          # 'MiR in protective stop. Wait'
          $ 1336 "AMR_Done≔ True "
          global AMR_Done=  True
        else:
          $ 1337 "ElseIf MiR_State≟3"
          if (modbus_get_signal_status("MiR_State") == 3):
            $ 1338 "AMR_Done≔ True "
            global AMR_Done=  True
          end
        end
      end
    elif (6 == switch_1):
      $ 1339 "Case 6"
      $ 1340 "execute"
      $ 1341 "AMR_AtTarget≔(AMR_PosActual≟AMR_PosTarget)"
      global AMR_AtTarget=(AMR_PosActual == AMR_PosTarget)
      $ 1342 "Switch AMR_Step"
      switch_2 = AMR_Step
      $ 1343 "Case 0"
      if (0 == switch_2):
        $ 1344 "If  not AMR_AtTarget"
        if (  not  AMR_AtTarget):
          $ 1345 "AMR_Step≔1"
          global AMR_Step=1
        else:
          $ 1346 "Else" "noBreak"
          $ 1347 "AMR_Done≔ True "
          global AMR_Done=  True
        end
      elif (1 == switch_2):
        $ 1348 "Case 1"
        $ 1349 "general Settings"
        $ 1350 "Set O2T_Acknowledge=0"
        modbus_set_output_register("O2T_Acknowledge", 0)
        $ 1351 "check for error"
        $ 1352 "If OBJ_Picked and MiR_State≟10"
        if (OBJ_Picked  and  modbus_get_signal_status("MiR_State") == 10):
          $ 1353 "Error"
          $ 1354 "set_error(ERROR_ROBOT_ARM_NOT_IN_HOME_POSE)"
          set_error(ERROR_ROBOT_ARM_NOT_IN_HOME_POSE)
          $ 1355 "Action≔0"
          global Action=0
        else:
          $ 1356 "ElseIf  not found_in_list(AMR_PosTarget, AMR_TargetList)"
          if (  not  found_in_list(AMR_PosTarget, AMR_TargetList)):
            $ 1357 "Error"
            $ 1358 "set_error(ERROR_UNKNOWN_POSE)"
            set_error(ERROR_UNKNOWN_POSE)
            $ 1359 "Action≔0"
            global Action=0
          end
        end
        $ 1360 "If MiR_State≟3"
        if (modbus_get_signal_status("MiR_State") == 3):
          $ 1361 "Set MiR_CMD_Start=Off"
          modbus_set_output_signal("MiR_CMD_Start", False)
          $ 1362 "Switch Action"
          switch_3 = Action
          $ 1363 "Case 51"
          if (51 == switch_3):
            $ 1364 "Charge"
            $ 1365 "'trigger the charging mission'"
            # 'trigger the charging mission'
            $ 1366 "'target pos is predefined'"
            # 'target pos is predefined'
            $ 1367 "Set O2T_Footprint=0"
            modbus_set_output_register("O2T_Footprint", 0)
            $ 1368 "Set O2T_Action=1"
            modbus_set_output_register("O2T_Action", 1)
            $ 1369 "If MiR_Mis_Queue≟0"
            if (modbus_get_signal_status("MiR_Mis_Queue") == 0):
              $ 1370 "Set O2T_Mis_Charge=On"
              modbus_set_output_signal("O2T_Mis_Charge", True)
              $ 1371 "Wait MiR_Mis_Queue≥1"
              while (not(modbus_get_signal_status("MiR_Mis_Queue") >= 1)):
                sync()
              end
              $ 1372 "Set O2T_Mis_Charge=Off"
              modbus_set_output_signal("O2T_Mis_Charge", False)
            end
          elif (52 == switch_3):
            $ 1373 "Case 52"
            $ 1374 "Navigate"
            $ 1375 "'trigger the standard missoin'"
            # 'trigger the standard missoin'
            $ 1376 "Set O2T_Footprint=AMR_FootprintID"
            modbus_set_output_register("O2T_Footprint", AMR_FootprintID)
            $ 1377 "Set O2T_Target_Pos=AMR_PosTarget"
            modbus_set_output_register("O2T_Target_Pos", AMR_PosTarget)
            $ 1378 "Set O2T_Action=2"
            modbus_set_output_register("O2T_Action", 2)
            $ 1379 "If MiR_Mis_Queue≟0"
            if (modbus_get_signal_status("MiR_Mis_Queue") == 0):
              $ 1380 "Set O2T_Mis_Main=On"
              modbus_set_output_signal("O2T_Mis_Main", True)
              $ 1381 "Wait MiR_Mis_Queue≥1"
              while (not(modbus_get_signal_status("MiR_Mis_Queue") >= 1)):
                sync()
              end
              $ 1382 "Set O2T_Mis_Main=Off"
              modbus_set_output_signal("O2T_Mis_Main", False)
            end
          end
        else:
          $ 1383 "ElseIf MiR_State≟4"
          if (modbus_get_signal_status("MiR_State") == 4):
            $ 1384 "Set MiR_CMD_Start=On"
            modbus_set_output_signal("MiR_CMD_Start", True)
          else:
            $ 1385 "ElseIf MiR_State≟5"
            if (modbus_get_signal_status("MiR_State") == 5):
              $ 1386 "AMR_Step≔2"
              global AMR_Step=2
            else:
              $ 1387 "ElseIf MiR_State≟10"
              if (modbus_get_signal_status("MiR_State") == 10):
                $ 1388 "'AMR still in safeguard stop'"
                # 'AMR still in safeguard stop'
              end
            end
          end
        end
      elif (2 == switch_2):
        $ 1389 "Case 2"
        $ 1390 "acknowledge handshake"
        $ 1391 "If T2O_Done≟1 and O2T_Acknowledge≟0"
        if (modbus_get_signal_status("T2O_Done") == 1  and  modbus_get_signal_status("O2T_Acknowledge") == 0):
          $ 1392 "Set O2T_Acknowledge=1"
          modbus_set_output_register("O2T_Acknowledge", 1)
        else:
          $ 1393 "ElseIf T2O_Done≟0 and O2T_Acknowledge≟1"
          if (modbus_get_signal_status("T2O_Done") == 0  and  modbus_get_signal_status("O2T_Acknowledge") == 1):
            $ 1394 "Set O2T_Acknowledge=0"
            modbus_set_output_register("O2T_Acknowledge", 0)
            $ 1395 "AMR_AtTarget≔(AMR_PosActual≟AMR_PosTarget)"
            global AMR_AtTarget=(AMR_PosActual == AMR_PosTarget)
            $ 1396 "AMR_Done≔ True "
            global AMR_Done=  True
          end
        end
      end
      $ 1397 "translate errors"
      $ 1398 "If AMR_Done"
      if (AMR_Done):
        $ 1399 "Switch T2O_Error_ID"
        switch_2 = modbus_get_signal_status("T2O_Error_ID")
        $ 1400 "Case 2003"
        if (2003 == switch_2):
          $ 1401 "error"
          $ 1402 "set_error(ERROR_NOT_DOCKED)"
          set_error(ERROR_NOT_DOCKED)
        elif (2007 == switch_2):
          $ 1403 "Case 2007"
          $ 1404 "error"
          $ 1405 "set_error(ERROR_NOT_REACHABLE_TARGET)"
          set_error(ERROR_NOT_REACHABLE_TARGET)
        elif (2008 == switch_2):
          $ 1406 "Case 2008"
          $ 1407 "error"
          $ 1408 "set_error(ERROR_CHARGING_NOT_STARTED)"
          set_error(ERROR_CHARGING_NOT_STARTED)
        end
      end
    elif (7 == switch_1):
      $ 1409 "Case 7"
      $ 1410 "completing"
      $ 1411 "If MiR_Mis_Queue>0"
      if (modbus_get_signal_status("MiR_Mis_Queue")>0):
        $ 1412 "Set MiR_CMD_Abort=On"
        modbus_set_output_signal("MiR_CMD_Abort", True)
        $ 1413 "Wait MiR_Mis_Queue≟0"
        while (not(modbus_get_signal_status("MiR_Mis_Queue") == 0)):
          sync()
        end
        $ 1414 "Set MiR_CMD_Abort=Off"
        modbus_set_output_signal("MiR_CMD_Abort", False)
      end
      $ 1415 "If MiR_State≟3 or MiR_State≟10"
      if (modbus_get_signal_status("MiR_State") == 3  or  modbus_get_signal_status("MiR_State") == 10):
        $ 1416 "AMR_Done≔ True "
        global AMR_Done=  True
      end
    elif (9 == switch_1):
      $ 1417 "Case 9"
      $ 1418 "holding"
      $ 1419 "Set MiR_CMD_Abort=On"
      modbus_set_output_signal("MiR_CMD_Abort", True)
      $ 1420 "If MiR_State≟3 or MiR_State≟10"
      if (modbus_get_signal_status("MiR_State") == 3  or  modbus_get_signal_status("MiR_State") == 10):
        $ 1421 "Set MiR_CMD_Abort=Off"
        modbus_set_output_signal("MiR_CMD_Abort", False)
        $ 1422 "AMR_Done≔ True "
        global AMR_Done=  True
      end
    elif (11 == switch_1):
      $ 1423 "Case 11"
      $ 1424 "unholding"
      $ 1425 "Set MiR_CMD_Start=On"
      modbus_set_output_signal("MiR_CMD_Start", True)
      $ 1426 "If MiR_State≠4"
      if (modbus_get_signal_status("MiR_State") != 4):
        $ 1427 "Set MiR_CMD_Start=Off"
        modbus_set_output_signal("MiR_CMD_Start", False)
        $ 1428 "AMR_Step≔0"
        global AMR_Step=0
        $ 1429 "AMR_Done≔ True "
        global AMR_Done=  True
      end
    elif (12 == switch_1):
      $ 1430 "Case 12"
      $ 1431 "suspending"
      $ 1432 "'none'"
      # 'none'
    elif (14 == switch_1):
      $ 1433 "Case 14"
      $ 1434 "unsuspending"
      $ 1435 "'none'"
      # 'none'
    elif (15 == switch_1):
      $ 1436 "Case 15"
      $ 1437 "aborting"
      $ 1438 "Set MiR_CMD_Abort=On"
      modbus_set_output_signal("MiR_CMD_Abort", True)
      $ 1439 "Wait MiR_State≟3"
      while (not(modbus_get_signal_status("MiR_State") == 3)):
        sync()
      end
      $ 1440 "Set MiR_CMD_Abort=Off"
      modbus_set_output_signal("MiR_CMD_Abort", False)
    elif (17 == switch_1):
      $ 1441 "Case 17"
      $ 1442 "clearing"
      $ 1443 "If MiR_Error_ID≠0"
      if (modbus_get_signal_status("MiR_Error_ID") != 0):
        $ 1444 "Set MiR_CMD_Clear_E=On"
        modbus_set_output_signal("MiR_CMD_Clear_E", True)
        $ 1445 "Wait MiR_Error_ID≟0"
        while (not(modbus_get_signal_status("MiR_Error_ID") == 0)):
          sync()
        end
        $ 1446 "Set MiR_CMD_Clear_E=Off"
        modbus_set_output_signal("MiR_CMD_Clear_E", False)
      end
      $ 1447 "If MiR_Error_ID≟0"
      if (modbus_get_signal_status("MiR_Error_ID") == 0):
        $ 1448 "AMR_Done≔ True "
        global AMR_Done=  True
      end
    end
    $ 1449 "'=========='"
    # '=========='
    $ 1450 "PostSettings"
    $ 1451 "AMR_Position≔struct(position_identifier=T2O_Current_Pos, x1=MiR_Position_X1, x2=MiR_Position_X2, y1=MiR_Position_Y1, y2=MiR_Position_Y2, theta1=MiR_Theta_1, theta2=MiR_Theta_2) "
    global AMR_Position=struct(position_identifier=modbus_get_signal_status("T2O_Current_Pos"), x1=modbus_get_signal_status("MiR_Position_X1"), x2=modbus_get_signal_status("MiR_Position_X2"), y1=modbus_get_signal_status("MiR_Position_Y1"), y2=modbus_get_signal_status("MiR_Position_Y2"), theta1=modbus_get_signal_status("MiR_Theta_1"), theta2=modbus_get_signal_status("MiR_Theta_2"))
  end
  def Sub_Action_V4():
    $ 1452 "Sub_Action_V4" "noBreak"
    $ 1453 "PreSettings"
    $ 1454 "init poses"
    $ 1455 "PSE_A≔p[0,0,0,0,0,0]"
    global PSE_A=p[0,0,0,0,0,0]
    $ 1456 "PSE_A_H≔p[0,0,0,0,0,0]"
    global PSE_A_H=p[0,0,0,0,0,0]
    $ 1457 "PSE_T≔p[0,0,0,0,0,0]"
    global PSE_T=p[0,0,0,0,0,0]
    $ 1458 "PSE_T_H≔p[0,0,0,0,0,0]"
    global PSE_T_H=p[0,0,0,0,0,0]
    $ 1459 "PSE_G≔p[0,0,0,0,0,0]"
    global PSE_G=p[0,0,0,0,0,0]
    $ 1460 "PSE_G_H≔p[0,0,0,0,0,0]"
    global PSE_G_H=p[0,0,0,0,0,0]
    $ 1461 "PSE_R≔p[0,0,0,0,0,0]"
    global PSE_R=p[0,0,0,0,0,0]
    $ 1462 "PSE_R_H≔p[0,0,0,0,0,0]"
    global PSE_R_H=p[0,0,0,0,0,0]
    $ 1463 "JNT_Q≔[0,0,0,0,0,0]"
    global JNT_Q=[0,0,0,0,0,0]
    $ 1464 "JNT_S≔[0,0,0,0,0,0]"
    global JNT_S=[0,0,0,0,0,0]
    $ 1465 "Gripping parameters"
    $ 1466 "OBJ = find_object_by_type(OBJs, OBJ_Type)"
    OBJ = find_object_by_type(OBJs, OBJ_Type)
    $ 1467 "GRP_Open_Pos≔OBJ.dimension.diameter * 1000 + 6"
    global GRP_Open_Pos=OBJ.dimension.diameter * 1000 + 6
    $ 1468 "GRP_Offset≔OBJ.gripper_offset"
    global GRP_Offset=OBJ.gripper_offset
    $ 1469 "rq_set_force_norm(50)"
     rq_set_force_norm (50)
    $ 1470 "rq_set_speed_norm(50)"
     rq_set_speed_norm (50)
    $ 1471 "Switch ITM_ID"
    switch_1 = ITM_ID
    $ 1472 "Case 1"
    if (1 == switch_1):
      $ 1473 "uML"
      $ 1474 "JIG2 = find_object_by_type(JIGs, JIG)"
      JIG2 = find_object_by_type(JIGs, JIG)
      $ 1475 "JIG_Offset≔JIG2.jig_offset"
      global JIG_Offset=JIG2.jig_offset
      $ 1476 "Switch JIG"
      switch_2 = JIG
      $ 1477 "Case 1"
      if (1 == switch_2):
        $ 1478 "3FG"
        $ 1479 "define poses"
        $ 1480 "FRM_Reference≔ULM_3FG"
        global FRM_Reference=ULM_3FG
        $ 1481 "JNT_Q≔JNT_HOME"
        global JNT_Q=JNT_HOME
        $ 1482 "PSE_T≔pose_trans(GRP_Offset, JIG_Offset)"
        global PSE_T= pose_trans (GRP_Offset, JIG_Offset)
        $ 1483 "PSE_A≔pose_trans(PSE_T, p[0,0,0.100,0,0,0])"
        global PSE_A= pose_trans (PSE_T, p[0,0,0.100,0,0,0])
        $ 1484 "PSE_R≔pose_add(PSE_T, p[0,0,0.100,0,0,0])"
        global PSE_R= pose_add (PSE_T, p[0,0,0.100,0,0,0])
      elif (2 == switch_2):
        $ 1485 "Case 2"
        $ 1486 "Input"
        $ 1487 "'CHANGE THE REFERENCE TO THE FRAME TO MOVE IN'"
        # 'CHANGE THE REFERENCE TO THE FRAME TO MOVE IN'
        $ 1488 "define poses"
        $ 1489 "FRM_Reference≔ULM_Input"
        global FRM_Reference=ULM_Input
        $ 1490 "PSE_T≔pose_trans(pose_trans(get_pattern_pos_rectangle(OBJ_Nbr, 'X', [10,5], patternsize=[0.181,0.081]), GRP_Offset), JIG_Offset)"
        global PSE_T= pose_trans ( pose_trans (get_pattern_pos_rectangle(OBJ_Nbr, "X", [10,5], patternsize=[0.181,0.081]), GRP_Offset), JIG_Offset)
        $ 1491 "If Action≟1"
        if (Action == 1):
          $ 1492 "PSE_R≔pose_add(PSE_T, p[0,0,0.200,0,0,0])"
          global PSE_R= pose_add (PSE_T, p[0,0,0.200,0,0,0])
          $ 1493 "PSE_A≔pose_add(PSE_T, p[0,0,0.100,0,0,0])"
          global PSE_A= pose_add (PSE_T, p[0,0,0.100,0,0,0])
        else:
          $ 1494 "ElseIf Action≟2"
          if (Action == 2):
            $ 1495 "PSE_R≔pose_add(PSE_T, p[0,0,0.100,0,0,0])"
            global PSE_R= pose_add (PSE_T, p[0,0,0.100,0,0,0])
            $ 1496 "PSE_A≔pose_add(PSE_T, p[0,0,0.200,0,0,0])"
            global PSE_A= pose_add (PSE_T, p[0,0,0.200,0,0,0])
          end
        end
      elif (3 == switch_2):
        $ 1497 "Case 3"
        $ 1498 "Output"
        $ 1499 "'CHANGE THE REFERENCE TO THE FRAME TO MOVE IN'"
        # 'CHANGE THE REFERENCE TO THE FRAME TO MOVE IN'
        $ 1500 "define poses"
        $ 1501 "FRM_Reference≔ULM_Output"
        global FRM_Reference=ULM_Output
        $ 1502 "PSE_T≔pose_trans(pose_trans(get_pattern_pos_rectangle(OBJ_Nbr, 'X', [10,5], patternsize=[0.181,0.081]), GRP_Offset), JIG_Offset)"
        global PSE_T= pose_trans ( pose_trans (get_pattern_pos_rectangle(OBJ_Nbr, "X", [10,5], patternsize=[0.181,0.081]), GRP_Offset), JIG_Offset)
        $ 1504 "If Action≟1"
        if (Action == 1):
          $ 1505 "PSE_R≔pose_add(PSE_T, p[0,0,0.200,0,0,0])"
          global PSE_R= pose_add (PSE_T, p[0,0,0.200,0,0,0])
          $ 1506 "PSE_A≔pose_add(PSE_T, p[0,0,0.100,0,0,0])"
          global PSE_A= pose_add (PSE_T, p[0,0,0.100,0,0,0])
        else:
          $ 1507 "ElseIf Action≟2"
          if (Action == 2):
            $ 1508 "PSE_R≔pose_add(PSE_T, p[0,0,0.100,0,0,0])"
            global PSE_R= pose_add (PSE_T, p[0,0,0.100,0,0,0])
            $ 1509 "PSE_A≔pose_add(PSE_T, p[0,0,0.200,0,0,0])"
            global PSE_A= pose_add (PSE_T, p[0,0,0.200,0,0,0])
          end
        end
      elif (4 == switch_2):
        $ 1510 "Case 4"
        $ 1511 "jig centrifuge racks"
        $ 1512 "define poses"
        $ 1513 "FRM_Reference≔ULM_Cent_Racks"
        global FRM_Reference=ULM_Cent_Racks
        $ 1514 "PSE_T≔get_pattern_pos_rectangle(JIG_Slot, 'X', [4,1], patternsize=[0.291,0])"
        global PSE_T=get_pattern_pos_rectangle(JIG_Slot, "X", [4,1], patternsize=[0.291,0])
        $ 1515 "If OBJ_Nbr≠0"
        if (OBJ_Nbr != 0):
          $ 1516 "PSE_T≔pose_trans(pose_trans(PSE_T, get_pattern_pos_rectangle(OBJ_Nbr, 'X', [3,3], patternsize=[0.060,0.060])),p[-0.030, -0.030,0,0,0,3.927])"
          global PSE_T= pose_trans ( pose_trans (PSE_T, get_pattern_pos_rectangle(OBJ_Nbr, "X", [3,3], patternsize=[0.060,0.060])),p[-0.030, -0.030,0,0,0,3.927])
        end
        $ 1517 "PSE_T≔pose_trans(PSE_T, GRP_Offset)"
        global PSE_T= pose_trans (PSE_T, GRP_Offset)
        $ 1518 "If Action≟1"
        if (Action == 1):
          $ 1519 "PSE_R≔pose_add(PSE_T, p[0,0,0.200,0,0,0])"
          global PSE_R= pose_add (PSE_T, p[0,0,0.200,0,0,0])
          $ 1520 "PSE_A≔pose_add(PSE_T, p[0,0,0.100,0,0,0])"
          global PSE_A= pose_add (PSE_T, p[0,0,0.100,0,0,0])
        else:
          $ 1521 "ElseIf Action≟2"
          if (Action == 2):
            $ 1522 "PSE_R≔pose_add(PSE_T, p[0,0,0.100,0,0,0])"
            global PSE_R= pose_add (PSE_T, p[0,0,0.100,0,0,0])
            $ 1523 "PSE_A≔pose_add(PSE_T, p[0,0,0.200,0,0,0])"
            global PSE_A= pose_add (PSE_T, p[0,0,0.200,0,0,0])
          end
        end
      elif (6 == switch_2):
        $ 1524 "Case 6"
        $ 1525 "Caps bin"
        $ 1526 "define poses"
        $ 1527 "'Drop cap'"
        # 'Drop cap'
        $ 1528 "FRM_Reference=ULM_Cap_Bin"
        FRM_Reference=ULM_Cap_Bin
        $ 1529 "PSE_T≔pose_RPY2RotVec(p[0,0,0,0,0,0])"
        global PSE_T=pose_RPY2RotVec(p[0,0,0,0,0,0])
        $ 1530 "PSE_T_H≔pose_add(PSE_T, p[0,0,-0.011,0,0,0])"
        global PSE_T_H= pose_add (PSE_T, p[0,0,-0.011,0,0,0])
        $ 1531 "PSE_A≔pose_trans(PSE_T, p[0,0,0.1,0,0,0])"
        global PSE_A= pose_trans (PSE_T, p[0,0,0.1,0,0,0])
        $ 1532 "PSE_R_H≔pose_add(PSE_T, p[0,0,0.100,0,0,0])"
        global PSE_R_H= pose_add (PSE_T, p[0,0,0.100,0,0,0])
        $ 1533 "PSE_R≔pose_add(PSE_T, p[0,0,0.100,0,0,0])"
        global PSE_R= pose_add (PSE_T, p[0,0,0.100,0,0,0])
      elif (7 == switch_2):
        $ 1534 "Case 7"
        $ 1535 "Sarstedt"
        $ 1536 "'CHANGE THE REFERENCE TO THE FRAME TO MOVE IN'"
        # 'CHANGE THE REFERENCE TO THE FRAME TO MOVE IN'
        $ 1542 "If TASK.ID≟10"
        if (TASK.ID == 10):
          $ 1543 "Frame & Position Params"
          $ 1545 "FRM_Reference = CAM_LM_SSRack"
          FRM_Reference = CAM_LM_SSRack
          $ 1550 "PSE_T≔uLM_SS_PickPlc"
          global PSE_T=uLM_SS_PickPlc
          $ 1551 "PSE_A≔pose_trans(PSE_T, p[0,0,0.1,0,0,0])"
          global PSE_A= pose_trans (PSE_T, p[0,0,0.1,0,0,0])
          $ 1552 "PSE_R≔pose_add(PSE_T, p[0,0,0.1,0,0,0])"
          global PSE_R= pose_add (PSE_T, p[0,0,0.1,0,0,0])
        else:
          $ 1553 "ElseIf TASK.ID≟11"
          if (TASK.ID == 11):
            $ 1554 "FRM_Reference = ULM_SS_Jig"
            FRM_Reference = ULM_SS_Jig
            $ 1555 "PSE_T≔pose_RPY2RotVec(p[0,0,0,0,0,0])"
            global PSE_T=pose_RPY2RotVec(p[0,0,0,0,0,0])
            $ 1556 "PSE_T≔pose_trans(PSE_T, GRP_Offset)"
            global PSE_T=pose_trans(PSE_T, GRP_Offset)
            $ 1557 "PSE_A≔pose_trans(PSE_T, p[0,0,0.1,0,0,0])"
            global PSE_A= pose_trans (PSE_T, p[0,0,0.1,0,0,0])
            $ 1558 "PSE_R≔pose_add(PSE_T, p[0,0,0.2,0,0,0])"
            global PSE_R= pose_add (PSE_T, p[0,0,0.2,0,0,0])
          end
        end
      elif (8 == switch_2):
        $ 1559 "Case 8"
        $ 1560 "NoK"
        $ 1561 "define poses"
        $ 1562 "'NoK'"
        # 'NoK'
        $ 1563 "FRM_Reference=ULM_NoK"
        FRM_Reference=ULM_NoK
        $ 1564 "PSE_T≔pose_RPY2RotVec(p[0,0,0,0,0,0])"
        global PSE_T=pose_RPY2RotVec(p[0,0,0,0,0,0])
        $ 1565 "PSE_A≔pose_trans(PSE_T, p[0,0,0.1,0,0,0])"
        global PSE_A= pose_trans (PSE_T, p[0,0,0.1,0,0,0])
        $ 1566 "PSE_R≔pose_add(PSE_T, p[0,0,0.100,0,0,0])"
        global PSE_R= pose_add (PSE_T, p[0,0,0.100,0,0,0])
      elif (9 == switch_2):
        $ 1567 "Case 9"
        $ 1568 "Pick_bott_jig"
        $ 1569 "define poses"
        $ 1570 "'NoK'"
        # 'NoK'
        $ 1571 "FRM_Reference=ULM_bottle_pick_const"
        FRM_Reference=p[0.0,0.0,0.0,0.0,0.0,0.0]
        $ 1572 "PSE_T≔pose_RPY2RotVec(p[0,0,0,0,0,0])"
        global PSE_T=pose_RPY2RotVec(p[0,0,0,0,0,0])
        $ 1573 "PSE_A≔pose_trans(PSE_T, p[0,0,0.1,0,0,0])"
        global PSE_A= pose_trans (PSE_T, p[0,0,0.1,0,0,0])
        $ 1574 "PSE_R≔pose_add(PSE_T, p[0,0,0.100,0,0,0])"
        global PSE_R= pose_add (PSE_T, p[0,0,0.100,0,0,0])
      elif (10 == switch_2):
        $ 1575 "Case 10"
        $ 1576 "Place_bott_jig"
        $ 1577 "define poses"
        $ 1578 "'NoK'"
        # 'NoK'
        $ 1579 "FRM_Reference=ULM_bottle_plac_const"
        FRM_Reference=p[0.0,0.0,0.0,0.0,0.0,0.0]
        $ 1580 "PSE_T≔pose_RPY2RotVec(p[0,0,0,0,0,0])"
        global PSE_T=pose_RPY2RotVec(p[0,0,0,0,0,0])
        $ 1581 "PSE_A≔pose_trans(PSE_T, p[0,0,0.1,0,0,0])"
        global PSE_A= pose_trans (PSE_T, p[0,0,0.1,0,0,0])
        $ 1582 "PSE_R≔pose_add(PSE_T, p[0,0,0.100,0,0,0])"
        global PSE_R= pose_add (PSE_T, p[0,0,0.100,0,0,0])
      elif (11 == switch_2):
        $ 1583 "Case 11"
        $ 1584 "Place_bott_jig"
        $ 1585 "define poses"
        $ 1586 "'NoK'"
        # 'NoK'
        $ 1587 "FRM_Reference=shake"
        FRM_Reference=shake
        $ 1588 "PSE_T≔pose_RPY2RotVec(p[0,0,0,0,0,0])"
        global PSE_T=pose_RPY2RotVec(p[0,0,0,0,0,0])
        $ 1589 "PSE_A≔pose_trans(PSE_T, p[0,0,0,0,0,0])"
        global PSE_A= pose_trans (PSE_T, p[0,0,0,0,0,0])
        $ 1590 "PSE_R≔pose_add(PSE_T, p[0,0,0,0,0,0])"
        global PSE_R= pose_add (PSE_T, p[0,0,0,0,0,0])
      elif (12 == switch_2):
        $ 1591 "Case 12"
        $ 1592 "Pick_Vial_jig"
        $ 1593 "define poses"
        $ 1594 "'NoK'"
        # 'NoK'
        $ 1595 "FRM_Reference=shake"
        FRM_Reference=shake
        $ 1596 "PSE_T≔pose_RPY2RotVec(p[0,0,0,0,0,0])"
        global PSE_T=pose_RPY2RotVec(p[0,0,0,0,0,0])
        $ 1597 "PSE_A≔pose_trans(PSE_T, p[0,0,0,0,0,0])"
        global PSE_A= pose_trans (PSE_T, p[0,0,0,0,0,0])
        $ 1598 "PSE_R≔pose_add(PSE_T, p[0,0,0,0,0,0])"
        global PSE_R= pose_add (PSE_T, p[0,0,0,0,0,0])
      end
    elif (2 == switch_1):
      $ 1599 "Case 2"
      $ 1600 "Centrifuge"
      $ 1601 "'CHANGE THE REFERENCE TO THE FRAME TO MOVE IN'"
      # 'CHANGE THE REFERENCE TO THE FRAME TO MOVE IN'
      $ 1602 "define poses"
      $ 1603 "FRM_Reference≔FRM_Centrifuge"
      global FRM_Reference=FRM_Centrifuge
      $ 1604 "PSE_T≔GRP_Offset"
      global PSE_T=GRP_Offset
      $ 1605 "If Action≟8"
      if (Action == 8):
        $ 1606 "PSE_R≔pose_add(PSE_T, p[0,0,0.250,0,0,0])"
        global PSE_R= pose_add (PSE_T, p[0,0,0.250,0,0,0])
        $ 1607 "PSE_A≔pose_add(PSE_T, p[0,0,0.150,0,0,0])"
        global PSE_A= pose_add (PSE_T, p[0,0,0.150,0,0,0])
      else:
        $ 1608 "ElseIf Action≟7"
        if (Action == 7):
          $ 1609 "PSE_R≔pose_add(PSE_T, p[0,0,0.150,0,0,0])"
          global PSE_R= pose_add (PSE_T, p[0,0,0.150,0,0,0])
          $ 1610 "PSE_A≔pose_add(PSE_T, p[0,0,0.250,0,0,0])"
          global PSE_A= pose_add (PSE_T, p[0,0,0.250,0,0,0])
        end
      end
    elif (3 == switch_1):
      $ 1611 "Case 3"
      $ 1612 "Output"
      $ 1613 "'CHANGE THE REFERENCE TO THE FRAME TO MOVE IN'"
      # 'CHANGE THE REFERENCE TO THE FRAME TO MOVE IN'
      $ 1614 "define poses"
      $ 1615 "FRM_Reference≔Base_const"
      global FRM_Reference=p[0.0,0.0,0.0,0.0,0.0,0.0]
      $ 1616 "PSE_T≔p[0,0,0,0,0,0]"
      global PSE_T=p[0,0,0,0,0,0]
      $ 1617 "PSE_A≔pose_add(PSE_T, p[0,0,0.150,0,0,0])"
      global PSE_A= pose_add (PSE_T, p[0,0,0.150,0,0,0])
      $ 1618 "PSE_R≔pose_add(PSE_T, p[0,0,0.100,0,0,0])"
      global PSE_R= pose_add (PSE_T, p[0,0,0.100,0,0,0])
    elif (5 == switch_1):
      $ 1619 "Case 5"
      $ 1620 "Sarstedt Pickup Table"
      $ 1621 "'CHANGE THE REFERENCE TO THE FRAME TO MOVE IN'"
      # 'CHANGE THE REFERENCE TO THE FRAME TO MOVE IN'
      $ 1622 "Switch JIG"
      switch_2 = JIG
      $ 1623 "Case 7"
      if (7 == switch_2):
        $ 1636 "Sarstedt"
        $ 1637 "'CHANGE THE REFERENCE TO THE FRAME TO MOVE IN'"
        # 'CHANGE THE REFERENCE TO THE FRAME TO MOVE IN'
        $ 1643 "If TASK.ID≟10"
        if (TASK.ID == 10):
          $ 1644 "Frame & Position Params"
          $ 1645 "FRM_Reference = CAM_LM_SSRack"
          FRM_Reference = CAM_LM_SSRack
          $ 1646 "PSE_T≔uLM_SS_PickPlc"
          global PSE_T=uLM_SS_PickPlc
          $ 1647 "PSE_A≔pose_trans(PSE_T, p[0,0,0.1,0,0,0])"
          global PSE_A= pose_trans (PSE_T, p[0,0,0.1,0,0,0])
          $ 1648 "PSE_R≔pose_add(PSE_T, p[0,0,0.1,0,0,0])"
          global PSE_R= pose_add (PSE_T, p[0,0,0.1,0,0,0])
        end
      end
    elif (13 == switch_1):
      $ 1655 "Case 13"
      $ 1656 "Sarstedt Pickup Table"
      $ 1657 "'CHANGE THE REFERENCE TO THE FRAME TO MOVE IN'"
      # 'CHANGE THE REFERENCE TO THE FRAME TO MOVE IN'
      $ 1658 "Switch JIG"
      switch_2 = JIG
      $ 1659 "Case 7"
      if (7 == switch_2):
        $ 1672 "Bottle"
        $ 1673 "'CHANGE THE REFERENCE TO THE FRAME TO MOVE IN'"
        # 'CHANGE THE REFERENCE TO THE FRAME TO MOVE IN'
        $ 1679 "If TASK.ID≟43"
        if (TASK.ID == 43):
          $ 1680 "Frame & Position Params"
          $ 1682 "PSE_T≔uLM_SS_PickPlc"
          global PSE_T=uLM_SS_PickPlc
          $ 1683 "PSE_A≔pose_trans(PSE_T, p[0,0,0.1,0,0,0])"
          global PSE_A= pose_trans (PSE_T, p[0,0,0.1,0,0,0])
          $ 1684 "PSE_R≔pose_add(PSE_T, p[0,0,0.1,0,0,0])"
          global PSE_R= pose_add (PSE_T, p[0,0,0.1,0,0,0])
        end
      end
    end
    $ 1691 "Additional check"
    $ 1692 "If  not is_reachable(FRM_Reference,[PSE_A,PSE_A_H,PSE_T,PSE_T_H,PSE_R,PSE_R_H])"
    if (  not  is_reachable(FRM_Reference,[PSE_A,PSE_A_H,PSE_T,PSE_T_H,PSE_R,PSE_R_H])):
      $ 1693 "Error"
      $ 1694 "set_error(ERROR_POSE_NOT_REACHABLE)"
      set_error(ERROR_POSE_NOT_REACHABLE)
      $ 1695 "Action≔0"
      global Action=0
    end
    $ 1696 "'=========='"
    # '=========='
    $ 1697 "Switch Action"
    switch_1 = Action
    $ 1698 "Case 1"
    if (1 == switch_1):
      $ 1699 "Pick"
      $ 1700 "Action_Info≔'pick object'"
      global Action_Info="pick object"
      $ 1701 "do_transition(pose_trans(FRM_Reference, PSE_T), keep_rxry=OBJ_Picked)"
      do_transition( pose_trans (FRM_Reference, PSE_T), keep_rxry=OBJ_Picked)
      $ 1702 "EOAT"
      $ 1703 "If  not OBJ_Picked"
      if (  not  OBJ_Picked):
        $ 1704 "rq_move_and_wait_mm(GRP_Open_Pos)"
         rq_move_and_wait_mm (GRP_Open_Pos)
      end
      $ 1705 "If PSE_A_H≠PSE_Z"
      if (PSE_A_H != PSE_Z):
        $ 1706 "If JNT_Q≠JNT_Z"
        if (JNT_Q != JNT_Z):
          $ 1707 "movej(get_inverse_kin(pose_trans(FRM_Reference, PSE_A_H), qnear=JNT_Q), r=0.050)"
          movej(get_inverse_kin( pose_trans (FRM_Reference, PSE_A_H), qnear=JNT_Q), r=0.050)
        else:
          $ 1708 "Else" "noBreak"
          $ 1709 "movej(pose_trans(FRM_Reference, PSE_A_H), r=0.050)"
          movej( pose_trans (FRM_Reference, PSE_A_H), r=0.050)
        end
      end
      $ 1710 "If PSE_A≠PSE_Z"
      if (PSE_A != PSE_Z):
        $ 1711 "If JNT_Q≠JNT_Z"
        if (JNT_Q != JNT_Z):
          $ 1712 "movej(get_inverse_kin(pose_trans(FRM_Reference, PSE_A), qnear=JNT_Q), r=0.020)"
          movej(get_inverse_kin( pose_trans (FRM_Reference, PSE_A), qnear=JNT_Q), r=0.020)
        else:
          $ 1713 "Else" "noBreak"
          $ 1714 "movej(pose_trans(FRM_Reference, PSE_A), r=0.020)"
          movej( pose_trans (FRM_Reference, PSE_A), r=0.020)
        end
      end
      $ 1715 "MoveL"
      $ 1716 "If PSE_T_H≠PSE_Z"
      if (PSE_T_H != PSE_Z):
        $ 1717 "PSE_T_H" "breakAfter"
        movel(pose_trans(FRM_Reference, PSE_T_H), a=0.5, v=0.4, r=0.01)
      end
      $ 1718 "PSE_T" "breakAfter"
      movel(pose_trans(FRM_Reference, PSE_T), a=0.08, v=0.12)
      $ 1719 "EOAT"
      $ 1720 "rq_set_force_norm(50)"
       rq_set_force_norm (50)
      $ 1721 "rq_close_and_wait()"
       rq_close_and_wait ()
      $ 1722 "OBJ_Picked≔rq_is_object_detected()"
      global OBJ_Picked= rq_is_object_detected ()
      $ 1723 "If  not OBJ_Picked"
      if (  not  OBJ_Picked):
        $ 1724 "set_error(ERROR_NO_OBJECT_TO_PICK)"
        set_error(ERROR_NO_OBJECT_TO_PICK)
      end
      $ 1725 "EXTT"
      $ 1726 "Switch JIG"
      switch_2 = JIG
      $ 1727 "Case 1"
      if (1 == switch_2):
        $ 1728 "3FG"
        $ 1729 "If OBJ_Picked"
        if (OBJ_Picked):
          $ 1730 "Set GRP_3F_Open=On"
          set_standard_digital_out(5, True)
        end
      end
      $ 1731 "If PSE_R_H≠PSE_Z"
      if (PSE_R_H != PSE_Z):
        $ 1732 "PSE_R" "breakAfter"
        movel(pose_trans(FRM_Reference, PSE_R), a=0.5, v=0.4, r=0.01)
        $ 1733 "PSE_R_H" "breakAfter"
        movel(pose_trans(FRM_Reference, PSE_R_H), a=0.5, v=0.4)
      else:
        $ 1734 "Else" "noBreak"
        $ 1735 "PSE_R" "breakAfter"
        movel(pose_trans(FRM_Reference, PSE_R), a=0.5, v=0.4)
      end
    elif (2 == switch_1):
      $ 1736 "Case 2"
      $ 1737 "Place"
      $ 1738 "Action_Info≔'place object'"
      global Action_Info="place object"
      $ 1739 "do_transition(pose_trans(FRM_Reference, PSE_T), keep_rxry=OBJ_Picked)"
      do_transition( pose_trans (FRM_Reference, PSE_T), keep_rxry=OBJ_Picked)
      $ 1740 "EXTT"
      $ 1741 "Switch JIG"
      switch_2 = JIG
      $ 1742 "Case 1"
      if (1 == switch_2):
        $ 1743 "3FG"
        $ 1744 "If OBJ_Picked"
        if (OBJ_Picked):
          $ 1745 "Set GRP_3F_Open=On"
          set_standard_digital_out(5, True)
        end
      end
      $ 1746 "If PSE_A_H≠PSE_Z"
      if (PSE_A_H != PSE_Z):
        $ 1747 "If JNT_Q≠JNT_Z"
        if (JNT_Q != JNT_Z):
          $ 1748 "movej(get_inverse_kin(pose_trans(FRM_Reference, PSE_A_H), qnear=JNT_Q), r=0.050)"
          movej(get_inverse_kin( pose_trans (FRM_Reference, PSE_A_H), qnear=JNT_Q), r=0.050)
        else:
          $ 1749 "Else" "noBreak"
          $ 1750 "movej(pose_trans(FRM_Reference, PSE_A_H), r=0.050)"
          movej( pose_trans (FRM_Reference, PSE_A_H), r=0.050)
        end
      end
      $ 1751 "If PSE_A≠PSE_Z"
      if (PSE_A != PSE_Z):
        $ 1752 "If JNT_Q≠JNT_Z"
        if (JNT_Q != JNT_Z):
          $ 1753 "movej(get_inverse_kin(pose_trans(FRM_Reference, PSE_A), qnear=JNT_Q), r=0.020)"
          movej(get_inverse_kin( pose_trans (FRM_Reference, PSE_A), qnear=JNT_Q), r=0.020)
        else:
          $ 1754 "Else" "noBreak"
          $ 1755 "movej(pose_trans(FRM_Reference, PSE_A), r=0.020)"
          movej( pose_trans (FRM_Reference, PSE_A), r=0.020)
        end
      end
      $ 1756 "MoveL"
      $ 1757 "If PSE_T_H≠PSE_Z"
      if (PSE_T_H != PSE_Z):
        $ 1758 "PSE_T_H" "breakAfter"
        movel(pose_trans(FRM_Reference, PSE_T_H), a=0.5, v=0.4, r=0.01)
      end
      $ 1759 "PSE_T" "breakAfter"
      global move_thread_flag_1759=0
      thread move_thread_1759():
        enter_critical
        move_thread_flag_1759 = 1
        movel(pose_trans(FRM_Reference, PSE_T), a=0.05, v=0.09)
        move_thread_flag_1759 = 2
        exit_critical
      end
      move_thread_flag_1759 = 0
      move_thread_han_1759 = run move_thread_1759()
      while (True):
        local targetTcpDirection=get_target_tcp_speed()
        local stepsToRetract=tool_contact(direction=targetTcpDirection)
        if (stepsToRetract > 0):
          kill move_thread_han_1759
          stopl(0.5)
          $ 1760 "Until (tool_contact_detection)"
          break
        end
        sleep(1.0E-10)
        if (move_thread_flag_1759 > 1):
          join move_thread_han_1759
          break
        end
        sync()
      end
      $ 1761 "Force"
      sleep(0.02)
      zero_ftsensor()
      force_mode(FRM_Reference, [1, 1, 1, 0, 0, 0], [0.0, 0.0, 0.0, 0.0, 0.0, 0.0], 2, [0.1, 0.1, 0.01, 0.3490658503988659, 0.3490658503988659, 0.3490658503988659])
      $ 1762 "PSE_T" "noBreak"
      movel(pose_trans(FRM_Reference, PSE_T), a=0.04, v=0.07)
      end_force_mode()
      stopl(5.0)
      $ 1763 "EXTT"
      $ 1764 "Switch JIG"
      switch_2 = JIG
      $ 1765 "Case 1"
      if (1 == switch_2):
        $ 1766 "3FG"
        $ 1767 "If OBJ_Picked"
        if (OBJ_Picked):
          $ 1768 "Set GRP_3F_Open=Off"
          set_standard_digital_out(5, False)
          $ 1769 "Wait: 0.2"
          sleep(0.2)
        end
      end
      $ 1770 "EOAT"
      $ 1771 "rq_move_and_wait_mm(GRP_Open_Pos)"
       rq_move_and_wait_mm (GRP_Open_Pos)
      $ 1772 "OBJ_Picked≔rq_is_object_detected()"
      global OBJ_Picked= rq_is_object_detected ()
      $ 1773 "If PSE_R_H≠PSE_Z"
      if (PSE_R_H != PSE_Z):
        $ 1774 "PSE_R" "breakAfter"
        movel(pose_trans(FRM_Reference, PSE_R), a=0.5, v=0.4, r=0.01)
        $ 1775 "PSE_R_H" "breakAfter"
        movel(pose_trans(FRM_Reference, PSE_R_H), a=0.5, v=0.4)
      else:
        $ 1776 "Else" "noBreak"
        $ 1777 "PSE_R" "breakAfter"
        movel(pose_trans(FRM_Reference, PSE_R), a=0.5, v=0.4)
      end
    elif (3 == switch_1):
      $ 1778 "Case 3"
      $ 1779 "Push"
      $ 1780 "Action_Info≔'push'"
      global Action_Info="push"
    elif (4 == switch_1):
      $ 1781 "Case 4"
      $ 1782 "Pull"
      $ 1783 "Action_Info≔'pull'"
      global Action_Info="pull"
    elif (6 == switch_1):
      $ 1786 "Case 6"
      $ 1787 "Drop the cap"
      $ 1788 "If JNT_A≠[0,0,0,0,0,0]"
      if (JNT_A != [0,0,0,0,0,0]):
        $ 1789 "MoveJ"
        $ 1790 "JNT_A" "breakAfter"
        movej(JNT_A, a=1.3962634015954636, v=1.7453292519943295, r=0.02)
      else:
        $ 1791 "Else" "noBreak"
        $ 1792 "MoveJ"
        $ 1793 "PSE_A" "breakAfter"
        movej(pose_trans(FRM_Reference, PSE_A), a=1.3962634015954636, v=1.7453292519943295, r=0.02)
      end
      $ 1794 "MoveL"
      $ 1795 "PSE_T" "breakAfter"
      movel(pose_trans(FRM_Reference, PSE_T), a=0.05, v=0.09)
      $ 1796 "'ADD OPEN GRIPPER'"
      # 'ADD OPEN GRIPPER'
      # begin: URCap Program Node
      #   Source: Robotiq_Grippers, 1.8.4.4844, Robotiq Inc.
      #   Type: Gripper
      $ 1797 "Gripper Move10mm (1)"
      if not(gripper_connected[0]):
        popup("Gripper 1 must be connected to run this program.", "No connection", False, True, True)
      end
      if not(rq_is_gripper_activated("1")):
        popup("Gripper 1 is not activated. Go to Installation tab > Gripper to activate it and run the program again.", "Not activated", False, True, True)
      end
      rq_set_pos_spd_for(201, 0, 28, "1")
      rq_wait_pos_spe_for_request(201, 0, 28, "1")
      rq_go_to("1")
      rq_wait("1")
      # end: URCap Program Node
      $ 1798 "PSE_T_H" "breakAfter"
      movel(pose_trans(FRM_Reference, PSE_T_H), a=0.05, v=0.09)
      # begin: URCap Program Node
      #   Source: Robotiq_Grippers, 1.8.4.4844, Robotiq Inc.
      #   Type: Gripper
      $ 1799 "Gripper Move40mm (1)"
      if not(gripper_connected[0]):
        popup("Gripper 1 must be connected to run this program.", "No connection", False, True, True)
      end
      if not(rq_is_gripper_activated("1")):
        popup("Gripper 1 is not activated. Go to Installation tab > Gripper to activate it and run the program again.", "Not activated", False, True, True)
      end
      rq_set_pos_spd_for(63, 0, 28, "1")
      rq_wait_pos_spe_for_request(63, 0, 28, "1")
      rq_go_to("1")
      rq_wait("1")
      # end: URCap Program Node
      $ 1800 "PSE_R" "breakAfter"
      movel(pose_trans(FRM_Reference, PSE_R), a=0.5, v=0.4)
    elif (7 == switch_1):
      $ 1801 "Case 7"
      $ 1802 "Load"
      $ 1803 "Action_Info≔'load object'"
      global Action_Info="load object"
      $ 1804 "do_transition(pose_trans(FRM_Reference, PSE_T), keep_rxry=OBJ_Picked)"
      do_transition( pose_trans (FRM_Reference, PSE_T), keep_rxry=OBJ_Picked)
      $ 1805 "If PSE_A_H≠PSE_Z"
      if (PSE_A_H != PSE_Z):
        $ 1806 "If JNT_Q≠JNT_Z"
        if (JNT_Q != JNT_Z):
          $ 1807 "movej(get_inverse_kin(pose_trans(FRM_Reference, PSE_A_H), qnear=JNT_Q), r=0.050)"
          movej(get_inverse_kin( pose_trans (FRM_Reference, PSE_A_H), qnear=JNT_Q), r=0.050)
        else:
          $ 1808 "Else" "noBreak"
          $ 1809 "movej(pose_trans(FRM_Reference, PSE_A_H), r=0.050)"
          movej( pose_trans (FRM_Reference, PSE_A_H), r=0.050)
        end
      end
      $ 1810 "If PSE_A≠PSE_Z"
      if (PSE_A != PSE_Z):
        $ 1811 "If JNT_Q≠JNT_Z"
        if (JNT_Q != JNT_Z):
          $ 1812 "movej(get_inverse_kin(pose_trans(FRM_Reference, PSE_A), qnear=JNT_Q), r=0.020)"
          movej(get_inverse_kin( pose_trans (FRM_Reference, PSE_A), qnear=JNT_Q), r=0.020)
        else:
          $ 1813 "Else" "noBreak"
          $ 1814 "movej(pose_trans(FRM_Reference, PSE_A), r=0.020)"
          movej( pose_trans (FRM_Reference, PSE_A), r=0.020)
        end
      end
      $ 1815 "MoveL"
      $ 1816 "If PSE_T_H≠PSE_Z"
      if (PSE_T_H != PSE_Z):
        $ 1817 "PSE_T_H" "breakAfter"
        movel(pose_trans(FRM_Reference, PSE_T_H), a=0.5, v=0.4, r=0.01)
      end
      $ 1818 "PSE_T" "breakAfter"
      global move_thread_flag_1818=0
      thread move_thread_1818():
        enter_critical
        move_thread_flag_1818 = 1
        movel(pose_trans(FRM_Reference, PSE_T), a=0.05, v=0.09)
        move_thread_flag_1818 = 2
        exit_critical
      end
      move_thread_flag_1818 = 0
      move_thread_han_1818 = run move_thread_1818()
      while (True):
        local targetTcpDirection=get_target_tcp_speed()
        local stepsToRetract=tool_contact(direction=targetTcpDirection)
        if (stepsToRetract > 0):
          kill move_thread_han_1818
          stopl(0.5)
          $ 1819 "Until (tool_contact_detection)"
          break
        end
        sleep(1.0E-10)
        if (move_thread_flag_1818 > 1):
          join move_thread_han_1818
          break
        end
        sync()
      end
      $ 1820 "Force"
      sleep(0.02)
      zero_ftsensor()
      force_mode(FRM_Reference, [0, 1, 1, 0, 0, 1], [0.0, 0.0, 0.0, 0.0, 0.0, 0.0], 2, [0.1, 0.05, 0.02, 0.3490658503988659, 0.3490658503988659, 3.141592653589793])
      $ 1821 "PSE_T" "noBreak"
      movel(pose_trans(FRM_Reference, PSE_T), a=0.04, v=0.07)
      end_force_mode()
      stopl(5.0)
      $ 1822 "EOAT"
      $ 1823 "rq_move_and_wait_mm(GRP_Open_Pos)"
       rq_move_and_wait_mm (GRP_Open_Pos)
      $ 1824 "OBJ_Picked≔rq_is_object_detected()"
      global OBJ_Picked= rq_is_object_detected ()
      $ 1825 "If PSE_R_H≠PSE_Z"
      if (PSE_R_H != PSE_Z):
        $ 1826 "PSE_R" "breakAfter"
        movel(pose_trans(FRM_Reference, PSE_R), a=0.5, v=0.4, r=0.01)
        $ 1827 "PSE_R_H" "breakAfter"
        movel(pose_trans(FRM_Reference, PSE_R_H), a=0.5, v=0.4)
      else:
        $ 1828 "Else" "noBreak"
        $ 1829 "PSE_R" "breakAfter"
        movel(pose_trans(FRM_Reference, PSE_R), a=0.5, v=0.4)
      end
    elif (8 == switch_1):
      $ 1830 "Case 8"
      $ 1831 "Unload"
      $ 1832 "Action_Info≔'pick object'"
      global Action_Info="pick object"
      $ 1833 "do_transition(pose_trans(FRM_Reference, PSE_T), keep_rxry=OBJ_Picked)"
      do_transition( pose_trans (FRM_Reference, PSE_T), keep_rxry=OBJ_Picked)
      $ 1834 "EOAT"
      $ 1835 "If  not OBJ_Picked"
      if (  not  OBJ_Picked):
        $ 1836 "rq_move_and_wait_mm(GRP_Open_Pos)"
         rq_move_and_wait_mm (GRP_Open_Pos)
      end
      $ 1837 "If PSE_A_H≠PSE_Z"
      if (PSE_A_H != PSE_Z):
        $ 1838 "If JNT_Q≠JNT_Z"
        if (JNT_Q != JNT_Z):
          $ 1839 "movej(get_inverse_kin(pose_trans(FRM_Reference, PSE_A_H), qnear=JNT_Q), r=0.050)"
          movej(get_inverse_kin( pose_trans (FRM_Reference, PSE_A_H), qnear=JNT_Q), r=0.050)
        else:
          $ 1840 "Else" "noBreak"
          $ 1841 "movej(pose_trans(FRM_Reference, PSE_A_H), r=0.050)"
          movej( pose_trans (FRM_Reference, PSE_A_H), r=0.050)
        end
      end
      $ 1842 "If PSE_A≠PSE_Z"
      if (PSE_A != PSE_Z):
        $ 1843 "If JNT_Q≠JNT_Z"
        if (JNT_Q != JNT_Z):
          $ 1844 "movej(get_inverse_kin(pose_trans(FRM_Reference, PSE_A), qnear=JNT_Q), r=0.020)"
          movej(get_inverse_kin( pose_trans (FRM_Reference, PSE_A), qnear=JNT_Q), r=0.020)
        else:
          $ 1845 "Else" "noBreak"
          $ 1846 "movej(pose_trans(FRM_Reference, PSE_A), r=0.020)"
          movej( pose_trans (FRM_Reference, PSE_A), r=0.020)
        end
      end
      $ 1847 "MoveL"
      $ 1848 "If PSE_T_H≠PSE_Z"
      if (PSE_T_H != PSE_Z):
        $ 1849 "PSE_T_H" "breakAfter"
        movel(pose_trans(FRM_Reference, PSE_T_H), a=0.5, v=0.4, r=0.01)
      end
      $ 1850 "PSE_T" "breakAfter"
      movel(pose_trans(FRM_Reference, PSE_T), a=0.08, v=0.12)
      $ 1851 "Force"
      sleep(0.02)
      zero_ftsensor()
      force_mode(FRM_Reference, [1, 1, 0, 0, 0, 0], [0.0, 0.0, 0.0, 0.0, 0.0, 0.0], 2, [0.05, 0.05, 0.1, 0.3490658503988659, 0.3490658503988659, 0.3490658503988659])
      $ 1852 "EOAT" "noBreak"
      $ 1853 "rq_set_force_norm(50)" "noBreak"
       rq_set_force_norm (50)
      $ 1854 "rq_close_and_wait()" "noBreak"
       rq_close_and_wait ()
      $ 1855 "OBJ_Picked≔rq_is_object_detected()" "noBreak"
      global OBJ_Picked= rq_is_object_detected ()
      $ 1856 "If  not OBJ_Picked" "noBreak"
      if (  not  OBJ_Picked):
        $ 1857 "set_error(ERROR_NO_OBJECT_TO_PICK)" "noBreak"
        set_error(ERROR_NO_OBJECT_TO_PICK)
      end
      $ 1858 "If PSE_R_H≠PSE_Z" "noBreak"
      if (PSE_R_H != PSE_Z):
        $ 1859 "PSE_R" "noBreak"
        movel(pose_trans(FRM_Reference, PSE_R), a=0.5, v=0.4, r=0.01)
        $ 1860 "PSE_R_H" "noBreak"
        movel(pose_trans(FRM_Reference, PSE_R_H), a=0.5, v=0.4)
      else:
        $ 1861 "Else" "noBreak"
        $ 1862 "PSE_R" "noBreak"
        movel(pose_trans(FRM_Reference, PSE_R), a=0.5, v=0.4)
      end
      end_force_mode()
      stopl(5.0)
    elif (11 == switch_1):
      $ 1863 "Case 11"
      $ 1864 "Place without opening gripper"
      $ 1865 "Action_Info≔'place object without gripper opening'"
      global Action_Info="place object without gripper opening"
      $ 1867 "movel(FRM_Container_S, a=0.025, v=0.015, r=0.00001)"
      movel(FRM_Container_S, a=0.025, v=0.015, r=0.00001)
      $ 1868 "EXTT"
      $ 1869 "Switch JIG"
      switch_2 = JIG
      $ 1870 "Case 1"
      if (1 == switch_2):
        $ 1871 "3FG"
        $ 1872 "If OBJ_Picked"
        if (OBJ_Picked):
          $ 1873 "Set GRP_3F_Open=On"
          set_standard_digital_out(5, True)
        end
      end
      $ 1874 "If PSE_A_H≠PSE_Z"
      if (PSE_A_H != PSE_Z):
        $ 1875 "If JNT_Q≠JNT_Z"
        if (JNT_Q != JNT_Z):
          $ 1876 "movej(get_inverse_kin(pose_trans(FRM_Reference, PSE_A_H), qnear=JNT_Q), r=0.050)"
          movej(get_inverse_kin( pose_trans (FRM_Reference, PSE_A_H), qnear=JNT_Q), r=0.050)
        else:
          $ 1877 "Else" "noBreak"
          $ 1878 "movej(pose_trans(FRM_Reference, PSE_A_H), r=0.050)"
          movej( pose_trans (FRM_Reference, PSE_A_H), r=0.050)
        end
      end
      $ 1879 "If PSE_A≠PSE_Z"
      if (PSE_A != PSE_Z):
        $ 1880 "If JNT_Q≠JNT_Z"
        if (JNT_Q != JNT_Z):
          $ 1881 "movej(get_inverse_kin(pose_trans(FRM_Reference, PSE_A), qnear=JNT_Q), r=0.020)"
          movej(get_inverse_kin( pose_trans (FRM_Reference, PSE_A), qnear=JNT_Q), r=0.020)
        else:
          $ 1882 "Else" "noBreak"
          $ 1883 "movej(pose_trans(FRM_Reference, PSE_A), r=0.020)"
          movej( pose_trans (FRM_Reference, PSE_A), r=0.020)
        end
      end
      $ 1884 "MoveL"
      $ 1885 "If PSE_T_H≠PSE_Z"
      if (PSE_T_H != PSE_Z):
        $ 1886 "PSE_T_H" "breakAfter"
        movel(pose_trans(FRM_Reference, PSE_T_H), a=0.5, v=0.4, r=0.01)
      end
      $ 1887 "PSE_T" "breakAfter"
      global move_thread_flag_1887=0
      thread move_thread_1887():
        enter_critical
        move_thread_flag_1887 = 1
        movel(pose_trans(FRM_Reference, PSE_T), a=0.05, v=0.09)
        move_thread_flag_1887 = 2
        exit_critical
      end
      move_thread_flag_1887 = 0
      move_thread_han_1887 = run move_thread_1887()
      while (True):
        local targetTcpDirection=get_target_tcp_speed()
        local stepsToRetract=tool_contact(direction=targetTcpDirection)
        if (stepsToRetract > 0):
          kill move_thread_han_1887
          stopl(0.5)
          $ 1888 "Until (tool_contact_detection)"
          break
        end
        sleep(1.0E-10)
        if (move_thread_flag_1887 > 1):
          join move_thread_han_1887
          break
        end
        sync()
      end
      $ 1889 "Force"
      sleep(0.02)
      zero_ftsensor()
      force_mode(FRM_Reference, [1, 1, 1, 0, 0, 0], [0.0, 0.0, 0.0, 0.0, 0.0, 0.0], 2, [0.1, 0.1, 0.01, 0.3490658503988659, 0.3490658503988659, 0.3490658503988659])
      $ 1890 "PSE_T" "noBreak"
      movel(pose_trans(FRM_Reference, PSE_T), a=0.04, v=0.07)
      end_force_mode()
      stopl(5.0)
      $ 1891 "EXTT"
      $ 1892 "Switch JIG"
      switch_2 = JIG
      $ 1893 "Case 1"
      if (1 == switch_2):
        $ 1894 "3FG"
        $ 1895 "If OBJ_Picked"
        if (OBJ_Picked):
          $ 1896 "Set GRP_3F_Open=Off"
          set_standard_digital_out(5, False)
          $ 1897 "Wait: 0.2"
          sleep(0.2)
        end
      end
      $ 1898 "EOAT"
      $ 1899 "Comment"
      # Comment
    elif (12 == switch_1):
      $ 1900 "Case 12"
      $ 1901 "Decap"
      $ 1902 "Action_Info≔'decapping'"
      global Action_Info="decapping"
      $ 1903 "Set GRP_3F_Enable=On"
      set_standard_digital_out(4, True)
      $ 1904 "Set GRP_3F_Decap=On"
      set_standard_digital_out(3, True)
      $ 1905 "Force"
      sleep(0.02)
      zero_ftsensor()
      force_mode(tool_pose(), [0, 0, 1, 0, 0, 0], [0.0, 0.0, 5.0, 0.0, 0.0, 0.0], 2, [0.1, 0.1, 0.15, 0.3490658503988659, 0.3490658503988659, 0.3490658503988659])
      $ 1906 "check_decapping(offset=0.015, timeout=5, abort=CMD_Hold)" "noBreak"
      check_decapping(offset=0.015, timeout=5, abort=CMD_Hold)
      end_force_mode()
      stopl(5.0)
      $ 1907 "Set GRP_3F_Decap=Off"
      set_standard_digital_out(3, False)
      $ 1908 "Set GRP_3F_Enable=Off"
      set_standard_digital_out(4, False)
      $ 1909 "MoveL"
      $ 1910 "PSE_R" "breakAfter"
      movel(pose_trans(FRM_Reference, PSE_R), a=0.8, v=0.15)
    elif (13 == switch_1):
      $ 1911 "Case 13"
      $ 1912 "TMR_Barcode: Reset"
      TMR_Barcode = 0
      $ 1913 "Read"
      $ 1914 "TMR_Barcode: Start"
      TMR_Barcode_is_counting = True
      $ 1915 "If TMR_Barcode<PRM_TO_Read_BC"
      global thread_flag_1915=0
      thread Thread_if_1915():
        $ 1916 "KeyenceTrigger"
        $ 1917 "Set OClearResult=HI:Pulse 0.2"
        thread SinglePulse22():
          write_output_boolean_register(2, True)
          sleep(0.2)
          write_output_boolean_register(2, False)
        end
        singlePulse22 = run SinglePulse22()
        $ 1918 "Wait: 0.5"
        sleep(0.5)
        $ 1919 "Set OTriggerBarcode=Off"
        write_output_boolean_register(1, False)
        $ 1920 "Wait: 0.5"
        sleep(0.5)
        $ 1921 "Set OTriggerBarcode=On"
        write_output_boolean_register(1, True)
        $ 1922 "Wait: 0.5"
        sleep(0.5)
        $ 1923 "Preorient"
        $ 1924 "TMR_Barcode: Reset"
        TMR_Barcode = 0
        $ 1925 "If ICmdExctd"
        if (read_input_boolean_register(12)):
          $ 1926 "Set GRP_3F_Decap=On"
          set_standard_digital_out(3, True)
          $ 1927 "Set GRP_3F_Enable=On"
          set_standard_digital_out(4, True)
          $ 1928 "Loop ICmdExctd"
          while (read_input_boolean_register(12)):
            $ 1929 "KeyenceTrigger"
            $ 1930 "Set OClearResult=HI:Pulse 0.1"
            thread SinglePulse23():
              write_output_boolean_register(2, True)
              sleep(0.1)
              write_output_boolean_register(2, False)
            end
            singlePulse23 = run SinglePulse23()
            $ 1931 "Wait: 0.3"
            sleep(0.3)
            $ 1932 "Set OTriggerBarcode=Off"
            write_output_boolean_register(1, False)
            $ 1933 "Wait: 0.3"
            sleep(0.3)
            $ 1934 "Set OTriggerBarcode=On"
            write_output_boolean_register(1, True)
            $ 1935 "Wait: 0.1"
            sleep(0.1)
          end
        end
        $ 1936 "If  not ICmdExctd"
        if (  not  read_input_boolean_register(12)):
          $ 1937 "Set GRP_3F_Decap=On"
          set_standard_digital_out(3, True)
          $ 1938 "Set GRP_3F_Enable=On"
          set_standard_digital_out(4, True)
          $ 1939 "Wait ICmdExctd=HI"
          while (read_input_boolean_register(12) == False):
            sync()
          end
        end
        $ 1940 "Set GRP_3F_Decap=Off"
        set_standard_digital_out(3, False)
        $ 1941 "Set GRP_3F_Enable=Off"
        set_standard_digital_out(4, False)
        $ 1942 "OBJ_Brc_OK≔ True "
        global OBJ_Brc_OK=  True
        thread_flag_1915 = 1
      end
      if (TMR_Barcode<PRM_TO_Read_BC):
        global thread_handler_1915=run Thread_if_1915()
        while (thread_flag_1915 == 0):
          if not(TMR_Barcode<PRM_TO_Read_BC):
            kill thread_handler_1915
            thread_flag_1915 = 2
          else:
            sync()
          end
        end
      else:
        thread_flag_1915 = 2
      end
      if (thread_flag_1915 == 2):
        $ 1943 "Else" "noBreak"
        $ 1944 "exeption"
        $ 1945 "error"
        $ 1947 "OBJ_Brc_OK≔ False "
        global OBJ_Brc_OK=  False
      end
      $ 1948 "Set GRP_3F_Decap=Off"
      set_standard_digital_out(3, False)
      $ 1949 "Set GRP_3F_Enable=Off"
      set_standard_digital_out(4, False)
      $ 1950 "Set OTriggerBarcode=Off"
      write_output_boolean_register(1, False)
    elif (15 == switch_1):
      $ 1951 "Case 15"
      $ 1952 "Detect"
      $ 1953 "Action_Info≔'detect'"
      global Action_Info="detect"
    elif (30 == switch_1):
      $ 1954 "Case 30"
      $ 1955 "Shake"
      $ 1956 "Action_Info≔'shake'"
      global Action_Info="shake"
      $ 1957 "do_transition(pose_trans(FRM_Reference, PSE_T), keep_rxry=OBJ_Picked)"
      do_transition( pose_trans (FRM_Reference, PSE_T), keep_rxry=OBJ_Picked)
      $ 1958 "If PSE_A_H≠PSE_Z"
      if (PSE_A_H != PSE_Z):
        $ 1959 "If JNT_Q≠JNT_Z"
        if (JNT_Q != JNT_Z):
          $ 1960 "movej(get_inverse_kin(pose_trans(FRM_Reference, PSE_A_H), qnear=JNT_Q), r=0.050)"
          movej(get_inverse_kin( pose_trans (FRM_Reference, PSE_A_H), qnear=JNT_Q), r=0.050)
        else:
          $ 1961 "Else" "noBreak"
          $ 1962 "movej(pose_trans(FRM_Reference, PSE_A_H), r=0.050)"
          movej( pose_trans (FRM_Reference, PSE_A_H), r=0.050)
        end
      end
      $ 1963 "If PSE_A≠PSE_Z"
      if (PSE_A != PSE_Z):
        $ 1964 "If JNT_Q≠JNT_Z"
        if (JNT_Q != JNT_Z):
          $ 1965 "movej(get_inverse_kin(pose_trans(FRM_Reference, PSE_A), qnear=JNT_Q), r=0.020)"
          movej(get_inverse_kin( pose_trans (FRM_Reference, PSE_A), qnear=JNT_Q), r=0.020)
        else:
          $ 1966 "Else" "noBreak"
          $ 1967 "movej(pose_trans(FRM_Reference, PSE_A), r=0.020)"
          movej( pose_trans (FRM_Reference, PSE_A), r=0.020)
        end
      end
      $ 1968 "MoveL"
      $ 1969 "If PSE_T_H≠PSE_Z"
      if (PSE_T_H != PSE_Z):
        $ 1970 "PSE_T_H" "breakAfter"
        movel(pose_trans(FRM_Reference, PSE_T_H), a=0.5, v=0.4, r=0.01)
      end
      $ 1971 "PSE_T" "breakAfter"
      movel(pose_trans(FRM_Reference, PSE_T), a=0.08, v=0.12)
      $ 1972 "EXTT"
      $ 1973 "Comment"
      # Comment
      $ 1974 "MoveJ"
      $ 1975 "Waypoint_6" "breakAfter"
      movej(get_inverse_kin(Waypoint_6_p, qnear=Waypoint_6_q), a=1.3962634015954636, v=1.0471975511965976)
      $ 1976 "MoveJ"
      $ 1977 "Waypoint_18" "breakAfter"
      movej(get_inverse_kin(Waypoint_18_p, qnear=Waypoint_18_q), a=1.3962634015954636, v=1.0471975511965976)
      $ 1978 "MoveJ"
      $ 1979 "Waypoint_12" "breakAfter"
      movej(get_inverse_kin(Waypoint_12_p, qnear=Waypoint_12_q), a=1.3962634015954636, v=1.0471975511965976)
      $ 1980 "MoveJ"
      $ 1981 "Waypoint_19" "breakAfter"
      movej(get_inverse_kin(Waypoint_19_p, qnear=Waypoint_19_q), a=1.3962634015954636, v=1.0471975511965976)
      $ 1982 "If PSE_R_H≠PSE_Z"
      if (PSE_R_H != PSE_Z):
        $ 1983 "PSE_R" "breakAfter"
        movel(pose_trans(FRM_Reference, PSE_R), a=0.5, v=0.4, r=0.01)
        $ 1984 "PSE_R_H" "breakAfter"
        movel(pose_trans(FRM_Reference, PSE_R_H), a=0.5, v=0.4)
      else:
        $ 1985 "Else" "noBreak"
        $ 1986 "PSE_R" "breakAfter"
        movel(pose_trans(FRM_Reference, PSE_R), a=0.5, v=0.4)
      end
    elif (31 == switch_1):
      $ 1987 "Case 31"
      $ 1988 "Action_Info≔'Pick_Vial'"
      global Action_Info="Pick_Vial"
      $ 1989 "Pick_Vial"
      # begin: URCap Program Node
      #   Source: Robotiq_Grippers, 1.8.4.4844, Robotiq Inc.
      #   Type: Gripper
      $ 1990 "Gripper Open (1)"
      if not(gripper_connected[0]):
        popup("Gripper 1 must be connected to run this program.", "No connection", False, True, True)
      end
      if not(rq_is_gripper_activated("1")):
        popup("Gripper 1 is not activated. Go to Installation tab > Gripper to activate it and run the program again.", "Not activated", False, True, True)
      end
      rq_set_pos_spd_for(0, 82, 71, "1")
      rq_wait_pos_spe_for_request(0, 82, 71, "1")
      rq_go_to("1")
      rq_wait("1")
      # end: URCap Program Node
      $ 1991 "MoveJ"
      $ 1992 "Vial_above" "breakAfter"
      movej(get_inverse_kin(Vial_above_p, qnear=Vial_above_q), a=0.5235987755982988, v=0.4363323129985824, r=0.05)
      $ 1993 "MoveL"
      $ 1994 "Vial_pick_point" "breakAfter"
      movel(Vial_pick_point_p, a=0.5, v=0.1)
      # begin: URCap Program Node
      #   Source: Robotiq_Grippers, 1.8.4.4844, Robotiq Inc.
      #   Type: Gripper
      $ 1995 "Gripper Close (1)"
      if not(gripper_connected[0]):
        popup("Gripper 1 must be connected to run this program.", "No connection", False, True, True)
      end
      if not(rq_is_gripper_activated("1")):
        popup("Gripper 1 is not activated. Go to Installation tab > Gripper to activate it and run the program again.", "Not activated", False, True, True)
      end
      rq_set_pos_spd_for(255, 71, 84, "1")
      rq_wait_pos_spe_for_request(255, 71, 84, "1")
      rq_go_to("1")
      rq_wait("1")
      # end: URCap Program Node
      $ 1996 "MoveL"
      $ 1997 "Waypoint_20" "breakAfter"
      movel(Waypoint_20_p, a=0.5, v=0.1, r=0.05)
      $ 1998 "Home (Safe)"
      movej([-1.2302089344500047, -1.2969853503591224, -1.875639182904262, -1.539621866126728, 1.5731943360401213, -2.80099559440227], a=1.3962634015954636, v=1.0471975511965976)
    elif (32 == switch_1):
      $ 1999 "Case 32"
      $ 2001 "decap_Vial"
      $ 2002 "Set GRP_3F_Open=On"
      set_standard_digital_out(5, True)
      $ 2003 "MoveJ"
      $ 2004 "Waypoint_33" "breakAfter"
      movej(get_inverse_kin(Waypoint_33_p, qnear=Waypoint_33_q), a=0.5235987755982988, v=0.4363323129985824)
      $ 2005 "MoveL"
      $ 2006 "Vial_3FG_place" "breakAfter"
      movel(Vial_3FG_place_p, a=0.5, v=0.1)
      $ 2007 "Set GRP_3F_Open=Off"
      set_standard_digital_out(5, False)
      $ 2008 "Wait: 0.5"
      sleep(0.5)
      $ 2009 "MoveL"
      $ 2010 "Waypoint_34" "breakAfter"
      movel(Waypoint_34_p, a=0.5, v=0.1, r=0.05)
      $ 2011 "MoveJ"
      $ 2012 "cap_dump" "breakAfter"
      movej(get_inverse_kin(cap_dump_p, qnear=cap_dump_q), a=0.5235987755982988, v=0.4363323129985824)
      # begin: URCap Program Node
      #   Source: Robotiq_Grippers, 1.8.4.4844, Robotiq Inc.
      #   Type: Gripper
      $ 2013 "Gripper Open (1)"
      if not(gripper_connected[0]):
        popup("Gripper 1 must be connected to run this program.", "No connection", False, True, True)
      end
      if not(rq_is_gripper_activated("1")):
        popup("Gripper 1 is not activated. Go to Installation tab > Gripper to activate it and run the program again.", "Not activated", False, True, True)
      end
      rq_set_pos_spd_for(0, 255, 255, "1")
      rq_wait_pos_spe_for_request(0, 255, 255, "1")
      rq_go_to("1")
      rq_wait("1")
      # end: URCap Program Node
      $ 2014 "MoveJ"
      $ 2015 "Waypoint_35" "breakAfter"
      movej(get_inverse_kin(Waypoint_35_p, qnear=Waypoint_35_q), a=0.5235987755982988, v=0.4363323129985824, r=0.05)
      $ 2016 "MoveL"
      $ 2017 "Vial_3FG_place" "breakAfter"
      movel(Vial_3FG_place_p, a=0.5, v=0.1)
      # begin: URCap Program Node
      #   Source: Robotiq_Grippers, 1.8.4.4844, Robotiq Inc.
      #   Type: Gripper
      $ 2018 "Gripper Close (1)"
      if not(gripper_connected[0]):
        popup("Gripper 1 must be connected to run this program.", "No connection", False, True, True)
      end
      if not(rq_is_gripper_activated("1")):
        popup("Gripper 1 is not activated. Go to Installation tab > Gripper to activate it and run the program again.", "Not activated", False, True, True)
      end
      rq_set_pos_spd_for(255, 204, 255, "1")
      rq_wait_pos_spe_for_request(255, 204, 255, "1")
      rq_go_to("1")
      rq_wait("1")
      # end: URCap Program Node
      $ 2025 "Decap"
      $ 2026 "Action_Info≔'decapping'"
      global Action_Info="decapping"
      $ 2027 "Set GRP_3F_Enable=On"
      set_standard_digital_out(4, True)
      $ 2028 "Set GRP_3F_Decap=On"
      set_standard_digital_out(3, True)
      $ 2029 "Force"
      sleep(0.02)
      zero_ftsensor()
      force_mode(p[0.0,0.0,0.0,0.0,0.0,0.0], [0, 0, 1, 0, 0, 0], [0.0, 0.0, 1.0, 0.0, 0.0, 0.0], 2, [0.1, 0.1, 0.001, 0.3490658503988659, 0.3490658503988659, 0.3490658503988659])
      $ 2030 "check_decapping(offset=0.015, timeout=10, abort=CMD_Hold)" "noBreak"
      check_decapping(offset=0.015, timeout=10, abort=CMD_Hold)
      end_force_mode()
      stopl(5.0)
      $ 2031 "Set GRP_3F_Decap=Off"
      set_standard_digital_out(3, False)
      $ 2032 "Set GRP_3F_Enable=Off"
      set_standard_digital_out(4, False)
      $ 2033 "MoveL"
      $ 2034 "Waypoint_36" "breakAfter"
      movel(Waypoint_36_p, a=0.5, v=0.1, r=0.05)
      $ 2035 "MoveJ"
      $ 2036 "cap_dump" "breakAfter"
      movej(get_inverse_kin(cap_dump_p, qnear=cap_dump_q), a=0.5235987755982988, v=0.4363323129985824)
      # begin: URCap Program Node
      #   Source: Robotiq_Grippers, 1.8.4.4844, Robotiq Inc.
      #   Type: Gripper
      $ 2037 "Gripper Open (1)"
      if not(gripper_connected[0]):
        popup("Gripper 1 must be connected to run this program.", "No connection", False, True, True)
      end
      if not(rq_is_gripper_activated("1")):
        popup("Gripper 1 is not activated. Go to Installation tab > Gripper to activate it and run the program again.", "Not activated", False, True, True)
      end
      rq_set_pos_spd_for(0, 204, 255, "1")
      rq_wait_pos_spe_for_request(0, 204, 255, "1")
      rq_go_to("1")
      rq_wait("1")
      # end: URCap Program Node
      $ 2038 "MoveJ"
      $ 2039 "Waypoint_37" "breakAfter"
      movej(get_inverse_kin(Waypoint_37_p, qnear=Waypoint_37_q), a=0.5235987755982988, v=0.4363323129985824, r=0.036)
    elif (33 == switch_1):
      $ 2040 "Case 33"
      $ 2041 "Shake and liquid transfer"
      $ 2042 "MoveL"
      $ 2043 "Vial_liq_above" "breakAfter"
      movel(Vial_liq_above_p, a=0.5, v=0.1)
      $ 2044 "Vial_liq_pick_1" "breakAfter"
      movel(Vial_liq_pick_1_p, a=0.5, v=0.1)
      $ 2045 "Vial_liq_pick_2" "breakAfter"
      movel(Vial_liq_pick_2_p, a=0.5, v=0.1)
      # begin: URCap Program Node
      #   Source: Robotiq_Grippers, 1.8.4.4844, Robotiq Inc.
      #   Type: Gripper
      $ 2046 "Gripper Close (1)"
      if not(gripper_connected[0]):
        popup("Gripper 1 must be connected to run this program.", "No connection", False, True, True)
      end
